FUNCTION "FRK_Release_DeclarationUnit" : Void
{ S7_Optimized_Access := 'TRUE' }
VERSION : 0.1
VAR_IN_OUT
    Unit : "FRK_Unit";
    Hal : "ST_DeclarationUnitHal";
END_VAR
BEGIN
    "FRK_UnitSetPermit"(Unit := #Unit, Ok := #Hal.Cell.Clamp.Permit, Diag := #Hal.Cell.Clamp.Diag);
END_FUNCTION
// Generated frame v0.24; change the declaration, then regenerate.
FUNCTION_BLOCK "FB_DeclarationUnit"
{ S7_Optimized_Access := 'TRUE' }
VERSION : 0.1
VAR_INPUT
    Execute {ExternalWritable := 'False'} : Bool;
    Abort {ExternalWritable := 'False'} : Bool;
    Command {ExternalWritable := 'False'} : DInt;
    ParCmd {ExternalWritable := 'False'} : "ST_DeclarationParCmd";
    ParentIndex {ExternalAccessible := 'False'; ExternalVisible := 'False'; ExternalWritable := 'False'} : DInt;
    Startup {ExternalAccessible := 'False'; ExternalVisible := 'False'; ExternalWritable := 'False'} : Bool;
END_VAR
VAR_OUTPUT
    Busy {ExternalWritable := 'False'} : Bool;
    Done {ExternalWritable := 'False'} : Bool;
    Error {ExternalWritable := 'False'} : Bool;
    Aborted {ExternalWritable := 'False'} : Bool;
    Held {ExternalWritable := 'False'} : Bool;
    ErrorID {ExternalWritable := 'False'} : DWord;
    Timing {ExternalWritable := 'False'} : "ST_ModuleTiming";
    OutCmd {ExternalWritable := 'False'} : "ST_DeclarationOutCmd";
END_VAR
VAR_IN_OUT
    Hal : "ST_DeclarationUnitHal";
END_VAR
VAR
    OutImm {ExternalWritable := 'False'} : "ST_UnitProbeImm";
    Status {ExternalWritable := 'False'} : "ST_ModuleStatus";
    Core {ExternalAccessible := 'False'; ExternalVisible := 'False'; ExternalWritable := 'False'} : "FRK_Core";
    Nameplate {ExternalWritable := 'False'} : "ST_Nameplate";
    EngineeringSlots {ExternalAccessible := 'False'; ExternalVisible := 'False'; ExternalWritable := 'False'} : Array[1..1] of Int;
    RunStyle {ExternalWritable := 'False'} : DInt;
    SupportedRunStylesPublished {ExternalWritable := 'False'} : Array[0..2] of Bool;
    HostEvents {ExternalWritable := 'False'} : "FRK_HostEvents";
    HostSeenSequence {ExternalAccessible := 'False'; ExternalVisible := 'False'; ExternalWritable := 'False'} : UDInt;
    HostDoneSeen {ExternalAccessible := 'False'; ExternalVisible := 'False'; ExternalWritable := 'False'} : Bool;
    SystemHealth {ExternalWritable := 'False'} : "ST_SystemHealthStatus";
    HealthBook {ExternalAccessible := 'False'; ExternalVisible := 'False'; ExternalWritable := 'False'} : "FRK_HealthBook";
    HealthConfig {ExternalAccessible := 'False'; ExternalVisible := 'False'; ExternalWritable := 'False'} : "ST_SystemHealthParCfg";
    SignalTower {ExternalWritable := 'False'} : "ST_SignalTowerOut";
    TowerBook {ExternalAccessible := 'False'; ExternalVisible := 'False'; ExternalWritable := 'False'} : "FRK_TowerBook";
    TowerConfig {ExternalAccessible := 'False'; ExternalVisible := 'False'; ExternalWritable := 'False'} : "ST_SignalTowerParCfg";
    ParCfg {ExternalWritable := 'False'} : "ST_ProductionUnitParCfg";
    LatchedParCmd {ExternalAccessible := 'False'; ExternalVisible := 'False'; ExternalWritable := 'False'} : "ST_DeclarationParCmd";
    StateFlags {ExternalWritable := 'False'} : Array[1..12] of "ST_StateFlag";
    StateFlagCount {ExternalWritable := 'False'} : Int;
    StateTouched {ExternalAccessible := 'False'; ExternalVisible := 'False'; ExternalWritable := 'False'} : Array[1..12] of Bool;
    Device {ExternalAccessible := 'False'; ExternalVisible := 'False'; ExternalWritable := 'False'} : "ST_UnitProbeDevice";
    StationCfg {ExternalWritable := 'False'} : "ST_UnitProbeStationCfg";
    ConfigStageParCfg {ExternalAccessible := 'False'; ExternalVisible := 'False'; ExternalWritable := 'False'} : "ST_ProductionUnitParCfg";
    ConfigDefaultParCfg {ExternalAccessible := 'False'; ExternalVisible := 'False'; ExternalWritable := 'False'} : "ST_ProductionUnitParCfg";
    ConfigStageStationCfg {ExternalAccessible := 'False'; ExternalVisible := 'False'; ExternalWritable := 'False'} : "ST_UnitProbeStationCfg";
    ConfigDefaultStationCfg {ExternalAccessible := 'False'; ExternalVisible := 'False'; ExternalWritable := 'False'} : "ST_UnitProbeStationCfg";
    ConfigStaged {ExternalAccessible := 'False'; ExternalVisible := 'False'; ExternalWritable := 'False'} : Bool;
    ConfigPersist {ExternalWritable := 'False'} : "ST_ConfigPersistStatus";
    Model {ExternalWritable := 'False'} : "ST_ModelId";
    AvailableModelCount {ExternalWritable := 'False'} : Int;
    AvailableModels {ExternalWritable := 'False'} : Array[1..3] of "ST_ModelId";
    ModelCapacity {ExternalWritable := 'False'} : Int;
    ModelGenerationSeen {ExternalAccessible := 'False'; ExternalVisible := 'False'; ExternalWritable := 'False'} : UDInt;
    ConfigSets {ExternalWritable := 'False'} : Array[1..4] of "ST_ConfigSetInfo";
    ConfigSetCount {ExternalWritable := 'False'} : Int;
    ConfigSetDocument {ExternalWritable := 'False'} : WString[480];
    ConfigSetDocumentLine {ExternalWritable := 'False'} : Int;
    ConfigSetDocumentLines {ExternalWritable := 'False'} : Int;
    SequenceViewEnabled {ExternalWritable := 'False'} : Bool;
    SequenceStepCount {ExternalWritable := 'False'} : Int;
    SequenceAnnotationCount {ExternalWritable := 'False'} : Int;
    Pending {ExternalWritable := 'False'} : "ST_Diagnostic";
    CurrentStep {ExternalWritable := 'False'} : "ST_StepRecord";
    CurrentStepElapsed {ExternalWritable := 'False'} : Time;
    CurrentStepTimedOut {ExternalWritable := 'False'} : Bool;
    SequenceSteps {ExternalWritable := 'False'} : Array[1..8] of "ST_SequenceStep";
    ActiveSteps {ExternalWritable := 'False'} : Array[0..0] of "ST_SequenceCursor";
    SequenceAnnotations {ExternalWritable := 'False'} : Array[1..4] of "ST_SequenceAnnotation";
    SequenceStepDef {ExternalAccessible := 'False'; ExternalVisible := 'False'; ExternalWritable := 'False'} : Array[1..8] of "ST_SequenceStepDef";
    Profiler {ExternalWritable := 'False'} : "FRK_Profiler_DeclarationUnit";
    Starved {ExternalWritable := 'False'} : Bool;
    Blocked {ExternalWritable := 'False'} : Bool;
    ProductionBook {ExternalAccessible := 'False'; ExternalVisible := 'False'; ExternalWritable := 'False'} : "FRK_Production";
    MachineState {ExternalWritable := 'False'} : DInt;
    Oee {ExternalWritable := 'False'} : "ST_Oee";
    OeeTrend {ExternalWritable := 'False'} : Array[1..60] of "ST_OeeSample";
    OeeTrendHead {ExternalWritable := 'False'} : Int;
    Unit {ExternalAccessible := 'False'; ExternalVisible := 'False'; ExternalWritable := 'False'} : "FRK_Unit";
    HmiRequest : "ST_HmiRequest";
    ModePolicy {ExternalAccessible := 'False'; ExternalVisible := 'False'; ExternalWritable := 'False'} : Array[0..6] of "ST_ModePolicy";
    Access {ExternalWritable := 'False'} : "FRK_Access";
    HmiResponse {ExternalWritable := 'False'} : "ST_HmiResponse";
    ConfigRev {ExternalWritable := 'False'} : UDInt;
    ConfigCursor {ExternalAccessible := 'False'; ExternalVisible := 'False'; ExternalWritable := 'False'} : "FRK_ConfigCursor";
    Part {ExternalWritable := 'False'} : "ST_PartContext";
    Decision {ExternalWritable := 'False'} : "ST_DecisionRequest";
    DecisionAnswer {ExternalWritable := 'False'} : Int;
    History {ExternalWritable := 'False'} : Array[1..16] of "ST_Diagnostic";
    HistoryHead {ExternalWritable := 'False'} : Int;
    AlarmLog {ExternalWritable := 'False'} : "FRK_AlarmLog";
    ModeActivePublished {ExternalWritable := 'False'} : DInt;
    RunningPublished {ExternalWritable := 'False'} : Bool;
    StopPendingPublished {ExternalWritable := 'False'} : Bool;
    SupportedModesPublished {ExternalWritable := 'False'} : Array[0..6] of Bool;
    GoodCount {ExternalWritable := 'False'} : UDInt;
    NokCount {ExternalWritable := 'False'} : UDInt;
    ReworkCount {ExternalWritable := 'False'} : UDInt;
    NokReason {ExternalWritable := 'False'} : DInt;
    Cell {ExternalWritable := 'False'} : "FB_DeclarationCell";
    Satellite {ExternalWritable := 'False'} : "FB_SatelliteUnit";
END_VAR
VAR_TEMP
    InstancePath : WString[254];
    RouteMatched : Bool;
    ManualMatched : Bool;
    ConfigRootIndex : Int;
    HealthResult : Bool;
END_VAR
VAR CONSTANT
    EXEC_READY : DInt := 0;
    MODULE_TIER : DInt := 1;
END_VAR
BEGIN
    // ---- GENERATED: setup
    IF #Startup OR NOT #Core.Named THEN
        #InstancePath := GetInstancePath(SIZE := 0);
        "FRK_SetIdentity"(Core := #Core, Status := #Status, InstancePath := #InstancePath,
            ModuleType := 1, TypeId := 1, Capabilities := DWORD#16#00000000, ParentIndex := #ParentIndex, TypeKey := 'Fraktal.Declaration.Unit');
        IF #Core.RegIndex = 1 THEN
            #Nameplate.ProductUri := WSTRING#'urn:fraktal:tia:operations:station-a';
            #Nameplate.ManufacturerName := 'Fraktal';
            #Nameplate.ProductDesignation := 'Isolated operations fixture';
        END_IF;
    END_IF;
    IF #Startup THEN "FRK_CfgRestore_DeclarationUnit"(Core := #Core, Status := #Status, ParCfg := #ParCfg, StationCfg := #StationCfg, ConfigStageParCfg := #ConfigStageParCfg, ConfigDefaultParCfg := #ConfigDefaultParCfg, ConfigStageStationCfg := #ConfigStageStationCfg, ConfigDefaultStationCfg := #ConfigDefaultStationCfg); END_IF;
    #ConfigRootIndex := "FRK_ConfigRoot"(RegIndex := #Core.RegIndex);
    "FRK_StateSweep"(Flags := #StateFlags, Count := #StateFlagCount, Touched := #StateTouched, Startup := #Startup);
    IF #Startup OR #ConfigRev = 0 THEN #ConfigRev := "FRK_ConfigRevision"(Previous := #ConfigRev); END_IF;
    #SupportedModesPublished[0] := TRUE;
    #SupportedModesPublished[1] := TRUE;
    #SupportedModesPublished[2] := TRUE;
    #SupportedModesPublished[3] := TRUE;
    #SupportedModesPublished[4] := FALSE;
    #SupportedModesPublished[5] := FALSE;
    #SupportedModesPublished[6] := FALSE;
    "FRK_UnitPrepare"(Core := #Core, Unit := #Unit, Policy := #ModePolicy, Request := #HmiRequest, Response := #HmiResponse, Startup := #Startup, InitialMode := 1);
    "FRK_AlarmBegin"(AlarmLog := #AlarmLog, Startup := #Startup);
    "FRK_AlarmHistoryBoot"(AlarmLog := #AlarmLog, Startup := #Startup, Scope := #Status.Name);
    "FRK_AlarmRecoveryBoot"(AlarmLog := #AlarmLog, Startup := #Startup, Scope := #Status.Name);
    "FRK_AlarmRecoveryTick"(AlarmLog := #AlarmLog);
    "FRK_AccessPolicyBoot"(Access := #Access, Startup := #Startup, Root := #Core.ParentIndex = 0, Scope := #Status.Name);
    "FRK_ClassBoot"(Access := #Access, Startup := #Startup, Root := #Core.ParentIndex = 0, Scope := #Status.Name);
    "FRK_AccessCyclic"(Access := #Access, Startup := #Startup, SourcePath := STRING_TO_WSTRING(#Status.Name), AlarmLog := #AlarmLog, Revision := #ConfigRev);
    "FRK_UnitMailbox"(Core := #Core, Unit := #Unit, Status := #Status, Policy := #ModePolicy, Access := #Access, Request := #HmiRequest, Response := #HmiResponse, Supported := #SupportedModesPublished);
    "FRK_ConfigStatus"(RootIndex := #ConfigRootIndex, Scope := #Status.Name, PolicyLost := (#Access.PolicyLost OR #Access.ClassesLost), UsersLost := "FRK_AccessStorage".UsersLost, Persist := #ConfigPersist, AlarmLog := #AlarmLog);
    #Unit.ConfigEnabled := #Core.ParentIndex = 0;
    #Unit.ConfigSetsEnabled := TRUE AND #Core.ParentIndex = 0;
    #Unit.ModelEnabled := #AvailableModelCount > 0;
    #Unit.ConfigBlocked := #ConfigPersist.RestoreLost AND NOT #ConfigPersist.RestoreAcknowledged AND #ConfigPersist.RestorePolicy = 1;
    #Unit.ConfigBlocked := #Unit.ConfigBlocked OR (#Access.PolicyLost OR #Access.ClassesLost);
    // ---- GENERATED: begin
    "FRK_Begin"(Core := #Core, Status := #Status, Execute := #Unit.RunReq, Abort := (#Abort OR #Unit.AbortReq), Command := 1);
    IF #Core.EvCommandStart THEN
        #LatchedParCmd := #ParCmd;
        CASE #Core.Command OF
            1: "FRK_UnitRunStart"(Core := #Core, Status := #Status, Timeout := #ParCfg.Timeout, Label := 'Run');
            ELSE "FRK_Start"(Core := #Core, Status := #Status, Supported := FALSE, Timeout := T#0ms, Label := '');
        END_CASE;
    END_IF;
    IF #Core.EvCommandStart THEN
    // ---- AUTHORED: CommandStart
    #Device.Received := "FRK_PartReceived"(Core := #Core, Unit := #Unit, Status := #Status, Part := #Part, AlarmLog := #AlarmLog);
    IF #Device.Received THEN
        "FRK_PartStarted"(Unit := #Unit, Status := #Status, Part := #Part, AlarmLog := #AlarmLog);
    END_IF;
    // ---- GENERATED: reaction end
    END_IF;
    IF #Core.EvCommandStart AND #Unit.Mode = 3 THEN
        "FRK_HostEmit"(Kind := 5, Scope := #Status.Name, PartUid := '', Subject := 'Model', Value := #Model.ModelCode, Verdict := 0, Reason := 0);
    END_IF;
    // ---- AUTHORED: cyclic management
    IF #Hal.Cell.Clamp.BackgroundFault THEN
        "FRK_Fault"(Core := #Core, Status := #Status, ReasonCode := 2901, Description := WSTRING#'test.unit.condition');
    END_IF;
    // ---- GENERATED: end management
    "FRK_Release_DeclarationUnit"(Unit := #Unit, Hal := #Hal);
    IF #Core.RegIndex > 0 THEN "FRK_Registry".Rows[#Core.RegIndex].AlarmBlocking := #AlarmLog.Blocking; END_IF;
    #Unit.AlarmBlocking := "FRK_AlarmTreeBlocking"(Owner := #Core.RegIndex) OR "FRK_AlarmRecoveryTreeBlocking"(Scope := #Status.Name);
    "FRK_UnitConsume"(Core := #Core, Unit := #Unit, Status := #Status, Policy := #ModePolicy, Access := #Access, Response := #HmiResponse, Supported := #SupportedModesPublished);
    "FRK_UnitMode"(Core := #Core, Unit := #Unit);
    #SupportedRunStylesPublished[0] := TRUE;
    #SupportedRunStylesPublished[1] := FALSE;
    #SupportedRunStylesPublished[2] := FALSE;
    "FRK_RunStylePrepare"(Owner := #Core.RegIndex, Startup := #Startup OR #Core.EvModeChanged OR #Unit.EvReset, Exec := #Core.Exec, Access := #Access, Supported := #SupportedRunStylesPublished);
    "FRK_RunStyleRequest"(Owner := #Core.RegIndex, Scope := #Status.Name, Exec := #Core.Exec, Supported := #SupportedRunStylesPublished, Unit := #Unit, Access := #Access, Response := #HmiResponse);
    "FRK_AlarmShelfRequest"(Scope := #Status.Name, Unit := #Unit, Access := #Access, Response := #HmiResponse, AlarmLog := #AlarmLog);
    #TowerConfig := "FRK_TowerDefaults".Config;
    "FRK_TowerRequest"(Scope := #Status.Name, Core := #Core, Unit := #Unit, Access := #Access, Response := #HmiResponse, Book := #TowerBook, ParCfg := #TowerConfig);
    "FRK_ProductionRequest"(Unit := #Unit, Access := #Access, Response := #HmiResponse, Book := #ProductionBook, Oee := #Oee, Trend := #OeeTrend, AlarmLog := #AlarmLog, Scope := #Status.Name);
    IF #Core.EvModeExit THEN
    // ---- AUTHORED: ModeExit
    #Device.ExitCalls := #Device.ExitCalls + 1;
    IF #Hal.Cell.Clamp.ExitHold THEN #Core.HookResult := 1; ELSE #Core.HookResult := 0; END_IF;
    // ---- GENERATED: reaction end
    END_IF;
    "FRK_UnitModeResolve"(Core := #Core, Unit := #Unit, Status := #Status, Policy := #ModePolicy, Timeout := #ParCfg.Timeout);
    IF #Core.EvModeChanged THEN
    // ---- AUTHORED: ModeChanged
    #Device.Changes := #Device.Changes + 1;
    // ---- GENERATED: reaction end
    END_IF;
    IF #Core.EvModeChanged THEN
        "FRK_HostEmit"(Kind := 9, Scope := #Status.Name, PartUid := '', Subject := 'Mode', Value := DINT_TO_STRING(#Unit.Mode), Verdict := 0, Reason := 0);
    END_IF;
    "FRK_SeqViewBegin"(Owner := #Core.RegIndex, Clear := #Startup OR #Core.EvModeChanged, ResetErrors := #Unit.EvReset, Enabled := #SequenceViewEnabled);
    "FRK_SeqProfilePrepare"(Owner := #Core.RegIndex, Run := #Core.Exec = 1 AND #Unit.Mode = 0, Withdraw := #Startup OR #Core.EvModeChanged);
    "FRK_DecisionCyclic"(Owner := #Core.RegIndex, Busy := #Core.Exec = 1, Reset := #Startup OR #Unit.EvReset OR #Core.EvModeChanged, AlarmLog := #AlarmLog);
    "FRK_UnitFollow"(Core := #Core, Unit := #Unit, Status := #Status, Policy := #ModePolicy, Access := #Access, Supported := #SupportedModesPublished);
    IF #Unit.RequestPending AND (#Unit.Request.Kind = 11 OR #Unit.Request.Kind = 16) THEN
        #ManualMatched := FALSE;
        #RouteMatched := "FRK_Route_DeclarationCell"(Module := #Cell, Hal := #Hal.Cell, Request := #Unit.Request, Report := #HmiResponse.Report);
        #ManualMatched := #ManualMatched OR #RouteMatched;
        #RouteMatched := "FRK_Route_SatelliteUnit"(Module := #Satellite, Hal := #Hal.Satellite, Request := #Unit.Request, Report := #HmiResponse.Report);
        #ManualMatched := #ManualMatched OR #RouteMatched;
        IF NOT #ManualMatched THEN
            "FRK_ReleaseReason"(Report := #HmiResponse.Report, Description := WSTRING#'std.error.unsupportedHmiRequest', Reason := 2008, Path := #Unit.Request.TargetPath, Kind := 4);
        END_IF;
        #HmiResponse.Accepted := #Unit.Request.Kind = 16 OR #HmiResponse.Report.Released;
        IF #Unit.Request.Kind = 11 THEN
            IF #HmiResponse.Accepted THEN #HmiResponse.Diagnostic := WSTRING#'std.audit.manualCommandAccepted'; ELSE #HmiResponse.Diagnostic := WSTRING#'std.audit.manualCommandRejected'; END_IF;
        END_IF;
    END_IF;
    IF #Unit.EvReset THEN "FRK_AlarmOperatorReset"(AlarmLog := #AlarmLog); END_IF;
    IF #Unit.EvReset THEN
    // ---- AUTHORED: OperatorReset
    #Device.Resets := #Device.Resets + 1;
    // ---- GENERATED: reset reaction end
    END_IF;
    IF #Core.ReleasePending OR #Unit.ReleaseChildren THEN
        "FRK_ReleaseCommand"(Core := #Cell.Core, Execute := #Cell.Execute);
        "FRK_ReleaseCommand"(Core := #Satellite.Core, Execute := #Satellite.Execute);
    END_IF;
    // ---- GENERATED: child call
    #Cell(ParentIndex := #Core.RegIndex, Startup := #Startup, Hal := #Hal.Cell);
    "FRK_ManualFinish"(Core := #Cell.Core, Execute := #Cell.Execute, ManualOwned := #Cell.ManualOwned);
    "FRK_UnitCascade"(ParentUnit := #Unit, Core := #Satellite.Core, Unit := #Satellite.Unit, Status := #Satellite.Status, Policy := #Satellite.ModePolicy, Access := #Satellite.Access, Supported := #Satellite.SupportedModesPublished, AlarmLog := #AlarmLog);
    // ---- GENERATED: child call
    #Satellite(ParentIndex := #Core.RegIndex, Startup := #Startup, Hal := #Hal.Satellite);
    #Unit.CascadePending := FALSE;
    "FRK_ConfigScratch".AccessRejected := FALSE;
    "FRK_CfgModelOperation_DeclarationUnit"(Core := #Core, Status := #Status, ParCfg := #ParCfg, Access := #Access, Unit := #Unit, HmiResponse := #HmiResponse, AlarmLog := #AlarmLog, ConfigPersist := #ConfigPersist, ConfigRev := #ConfigRev, AvailableModelCount := #AvailableModelCount, ModelCapacity := #ModelCapacity, ModelGenerationSeen := #ModelGenerationSeen, AvailableModels := #AvailableModels, StationCfg := #StationCfg, ConfigStageParCfg := #ConfigStageParCfg, ConfigStageStationCfg := #ConfigStageStationCfg, Cell := #Cell, Satellite := #Satellite);
    "FRK_CfgOperation_DeclarationUnit"(Core := #Core, Status := #Status, OutImm := #OutImm, ParCfg := #ParCfg, ModePolicy := #ModePolicy, Access := #Access, Unit := #Unit, HmiResponse := #HmiResponse, AlarmLog := #AlarmLog, ConfigPersist := #ConfigPersist, ConfigCursor := #ConfigCursor, ConfigRev := #ConfigRev, Model := #Model, AvailableModelCount := #AvailableModelCount, ConfigStaged := #ConfigStaged, ModelCapacity := #ModelCapacity, SequenceStepDef := #SequenceStepDef, SequenceStepCount := #SequenceStepCount, SupportedModesPublished := #SupportedModesPublished, StationCfg := #StationCfg, ConfigStageParCfg := #ConfigStageParCfg, ConfigDefaultParCfg := #ConfigDefaultParCfg, Cell := #Cell, Satellite := #Satellite);
    "FRK_CfgSetOperation_DeclarationUnit"(Core := #Core, Status := #Status, ParCfg := #ParCfg, ModePolicy := #ModePolicy, Access := #Access, Unit := #Unit, HmiResponse := #HmiResponse, ConfigPersist := #ConfigPersist, ConfigRev := #ConfigRev, Model := #Model, AvailableModelCount := #AvailableModelCount, ConfigSets := #ConfigSets, ConfigSetCount := #ConfigSetCount, ConfigSetDocument := #ConfigSetDocument, ConfigSetDocumentLine := #ConfigSetDocumentLine, ConfigSetDocumentLines := #ConfigSetDocumentLines, SupportedModesPublished := #SupportedModesPublished, StationCfg := #StationCfg, ConfigStageParCfg := #ConfigStageParCfg, ConfigStageStationCfg := #ConfigStageStationCfg, Cell := #Cell, Satellite := #Satellite, Startup := #Startup);
    IF #Unit.RequestPending AND #Core.ParentIndex = 0 THEN "FRK_SetResult"(Request := #Unit.Request, Response := #HmiResponse, Persist := #ConfigPersist, AlarmLog := #AlarmLog, Scope := #Status.Name, RootIndex := #ConfigRootIndex); END_IF;
    "FRK_ConfigAccessRefusal"(Unit := #Unit, Access := #Access, Response := #HmiResponse, Persist := #ConfigPersist, AlarmLog := #AlarmLog);
    "FRK_ConfigStatus"(RootIndex := #ConfigRootIndex, Scope := #Status.Name, PolicyLost := (#Access.PolicyLost OR #Access.ClassesLost), UsersLost := "FRK_AccessStorage".UsersLost, Persist := #ConfigPersist, AlarmLog := #AlarmLog);
    "FRK_RouteAbort"(Core := #Core, Abort := (#Abort OR #Unit.AbortReq));
    IF #Core.EvAbort THEN
        "FRK_PartAborted"(Core := #Core, Unit := #Unit, Status := #Status, Part := #Part, AlarmLog := #AlarmLog);
    END_IF;
    "FRK_SeqLifecycleUpdate"(Owner := #Core.RegIndex, Exec := #Core.Exec, Restart := #Startup OR #Core.EvModeChanged OR #Core.EvAbortInError);
    "FRK_DiagComposite"(Core := #Core, Status := #Status, AdoptErrors := FALSE);
    IF #Core.Dispatch AND #Core.RegIndex > 0 AND NOT "FRK_Registry".Fault THEN
    // ---- AUTHORED: dispatch
    IF #Hal.Cell.Clamp.Finish THEN
        #Device.Processed := FALSE;
        IF #Unit.CarrierIndex = 0 THEN
            #Device.Processed := TRUE;
        ELSE
            #Device.Processed := "FRK_PartProcessed"(Core := #Core, Unit := #Unit, Status := #Status, Part := #Part, AlarmLog := #AlarmLog, Verdict := #Hal.Cell.Clamp.Verdict, Reason := #Hal.Cell.Clamp.Diag.ReasonCode);
        END_IF;
        IF #Device.Processed THEN
            #Device.Cycles := #Device.Cycles + 1;
            IF #Unit.StopReq THEN
                "FRK_Complete"(Core := #Core, Status := #Status);
            ELSE
                #Device.Received := "FRK_PartReceived"(Core := #Core, Unit := #Unit, Status := #Status, Part := #Part, AlarmLog := #AlarmLog);
                IF #Device.Received THEN
                    "FRK_PartStarted"(Unit := #Unit, Status := #Status, Part := #Part, AlarmLog := #AlarmLog);
                END_IF;
            END_IF;
        END_IF;
    END_IF;
    // ---- GENERATED: end dispatch
    END_IF;
    "FRK_SeqViewEnd"(Owner := #Core.RegIndex, Revision := #ConfigRev, Fallback := #ParCfg.Timeout);
    "FRK_SeqViewDiagnostic"(Owner := #Core.RegIndex, Core := #Core, Status := #Status, Pending := #Pending);
    CASE #Core.RegIndex OF
        1:
            #SequenceStepDef := "FRK_Views".V001.Defs;
            #SequenceSteps := "FRK_Views".V001.Rows;
            #ActiveSteps := "FRK_Views".V001.Cursors;
            #SequenceAnnotations := "FRK_Views".V001.Notes;
            #SequenceStepCount := "FRK_Views".V001.Count;
            #SequenceAnnotationCount := "FRK_Views".V001.NoteCount;
            #CurrentStep := "FRK_Views".V001.Current;
            #CurrentStepElapsed := "FRK_Views".V001.Cursors[0].Elapsed;
            #CurrentStepTimedOut := "FRK_Views".V001.Cursors[0].TimedOut;
        13:
            #SequenceStepDef := "FRK_Views".V013.Defs;
            #SequenceSteps := "FRK_Views".V013.Rows;
            #ActiveSteps := "FRK_Views".V013.Cursors;
            #SequenceAnnotations := "FRK_Views".V013.Notes;
            #SequenceStepCount := "FRK_Views".V013.Count;
            #SequenceAnnotationCount := "FRK_Views".V013.NoteCount;
            #CurrentStep := "FRK_Views".V013.Current;
            #CurrentStepElapsed := "FRK_Views".V013.Cursors[0].Elapsed;
            #CurrentStepTimedOut := "FRK_Views".V013.Cursors[0].TimedOut;
        ELSE #SequenceViewEnabled := FALSE;
    END_CASE;
    "FRK_End"(Core := #Core, Status := #Status,
        Busy => #Busy, Done => #Done, Error => #Error, Aborted => #Aborted, Held => #Held, ErrorID => #ErrorID, Timing => #Timing);
    "FRK_SeqLifecycleUpdate"(Owner := #Core.RegIndex, Exec := #Core.Exec, Restart := FALSE);
    IF #Core.Exec = 3 OR #Core.Exec = 4 THEN
        "FRK_SeqProfilePrepare"(Owner := #Core.RegIndex, Run := FALSE, Withdraw := TRUE);
    END_IF;
    "FRK_SeqProfileEnd"(Owner := #Core.RegIndex, StepNo := #CurrentStep.StepNo, Expected := #CurrentStep.ExpectedTime, NowMs := "FRK_Clock".NowMs);
    CASE #Core.RegIndex OF
        1:
            #Profiler.LastCycle.CycleNo := "FRK_Profiles".P001.Book.Last.CycleNo;
            #Profiler.LastCycle.Started := "FRK_Profiles".P001.Book.Last.Started;
            #Profiler.LastCycle.StartedTimeSynchronized := "FRK_Profiles".P001.Book.Last.StartedTimeSynchronized;
            #Profiler.LastCycle.Total := "FRK_Profiles".P001.Book.Last.Total;
            #Profiler.LastCycle.WorkTime := "FRK_Profiles".P001.Book.Last.WorkTime;
            #Profiler.LastCycle.WaitTime := "FRK_Profiles".P001.Book.Last.WaitTime;
            #Profiler.LastCycle.ByClass := "FRK_Profiles".P001.Book.Last.ByClass;
            #Profiler.LastCycle.NSteps := "FRK_Profiles".P001.Book.LastNSteps;
            #Profiler.LastCycle.Truncated := "FRK_Profiles".P001.Book.LastTruncated;
            #Profiler.LastCycle.Steps := "FRK_Profiles".P001.LastSteps;
            #Profiler.StepStats := "FRK_Profiles".P001.Stats;
            #Profiler.StatsTruncated := "FRK_Profiles".P001.Book.StatsTruncated;
            #Profiler.LastCycleTime := "FRK_Profiles".P001.Book.LastCycleTime;
            #Profiler.MinCycleTime := "FRK_Profiles".P001.Book.MinCycleTime;
            #Profiler.History := "FRK_Profiles".P001.History;
            #Profiler.HistoryHead := "FRK_Profiles".P001.Book.Head;
        13:
            #Profiler.LastCycle.CycleNo := "FRK_Profiles".P013.Book.Last.CycleNo;
            #Profiler.LastCycle.Started := "FRK_Profiles".P013.Book.Last.Started;
            #Profiler.LastCycle.StartedTimeSynchronized := "FRK_Profiles".P013.Book.Last.StartedTimeSynchronized;
            #Profiler.LastCycle.Total := "FRK_Profiles".P013.Book.Last.Total;
            #Profiler.LastCycle.WorkTime := "FRK_Profiles".P013.Book.Last.WorkTime;
            #Profiler.LastCycle.WaitTime := "FRK_Profiles".P013.Book.Last.WaitTime;
            #Profiler.LastCycle.ByClass := "FRK_Profiles".P013.Book.Last.ByClass;
            #Profiler.LastCycle.NSteps := "FRK_Profiles".P013.Book.LastNSteps;
            #Profiler.LastCycle.Truncated := "FRK_Profiles".P013.Book.LastTruncated;
            #Profiler.LastCycle.Steps := "FRK_Profiles".P013.LastSteps;
            #Profiler.StepStats := "FRK_Profiles".P013.Stats;
            #Profiler.StatsTruncated := "FRK_Profiles".P013.Book.StatsTruncated;
            #Profiler.LastCycleTime := "FRK_Profiles".P013.Book.LastCycleTime;
            #Profiler.MinCycleTime := "FRK_Profiles".P013.Book.MinCycleTime;
            #Profiler.History := "FRK_Profiles".P013.History;
            #Profiler.HistoryHead := "FRK_Profiles".P013.Book.Head;
        ELSE RETURN;
    END_CASE;
    #Starved := #Core.Exec = 1 AND #Unit.Mode = 0 AND #CurrentStep.TimeClass = 1;
    #Blocked := #Core.Exec = 1 AND #Unit.Mode = 0 AND #CurrentStep.TimeClass = 2;
    "FRK_DecisionCyclic"(Owner := #Core.RegIndex, Busy := #Core.Exec = 1, Reset := #Startup OR #Unit.EvReset OR #Core.EvModeChanged, AlarmLog := #AlarmLog);
    "FRK_DecisionPublish"(Owner := #Core.RegIndex, Decision := #Decision, DecisionAnswer := #DecisionAnswer);
    IF NOT #Unit.EvReset THEN
        "FRK_AlarmCapture"(AlarmLog := #AlarmLog, Core := #Core, Status := #Status);
        "FRK_Capture_DeclarationCell"(Module := #Cell, AlarmLog := #AlarmLog);
        "FRK_AlarmEnd"(AlarmLog := #AlarmLog);
    END_IF;
    IF #Core.RegIndex > 0 THEN "FRK_Registry".Rows[#Core.RegIndex].AlarmBlocking := #AlarmLog.Blocking; END_IF;
    #Unit.AlarmBlocking := "FRK_AlarmTreeBlocking"(Owner := #Core.RegIndex) OR "FRK_AlarmRecoveryTreeBlocking"(Scope := #Status.Name);
    "FRK_ClassOperation"(Access := #Access, Unit := #Unit, Response := #HmiResponse, Scope := #Status.Name);
    "FRK_AccessPersist"(Access := #Access, Unit := #Unit, Response := #HmiResponse, SourcePath := STRING_TO_WSTRING(#Status.Name), AlarmLog := #AlarmLog);
    IF #Core.ParentIndex = 0 THEN "FRK_EngineeringTick"(Scope := #Status.Name, Slots := #EngineeringSlots, AlarmLog := #AlarmLog); END_IF;
    #HealthConfig := "FRK_HealthDefaults".Config;
    #HealthResult := "FRK_HealthCyclic"(Configured := TRUE, Scope := #Status.Name, Input := "FRK_HealthProbe".Input, ParCfg := #HealthConfig, Status := #SystemHealth, Book := #HealthBook, AlarmLog := #AlarmLog);
    IF #Startup THEN #ProductionBook := "FRK_ProductionDefaults".Book; #Oee := "FRK_ProductionDefaults".Oee; END_IF;
    #MachineState := "FRK_MachineState"(Exec := #Core.Exec, Mode := #Unit.Mode, Blocking := #Unit.AlarmBlocking, Starved := #Starved, Blocked := #Blocked, StopRequested := #Unit.StopReq);
    "FRK_OeeTick"(NowMs := "FRK_Clock".NowMs, Exec := #Core.Exec, Blocking := #Unit.AlarmBlocking, Good := #Unit.Good, Nok := #Unit.Nok, IdealCycleMs := #ParCfg.IdealCycleMs, Book := #ProductionBook, Oee := #Oee, Trend := #OeeTrend);
    #OeeTrendHead := #ProductionBook.TrendHead;
    IF "FRK_WorkDegradation"(CycleNo := #Profiler.LastCycle.CycleNo, WorkMs := TIME_TO_UDINT(#Profiler.LastCycle.WorkTime), BaselineMs := #ParCfg.BaselineMs, BandPercent := #StationCfg.DegradationPercent, Book := #ProductionBook) THEN
        "FRK_AlarmMessage"(AlarmLog := #AlarmLog, Reason := 2007, Description := WSTRING#'std.maintenance.cycleTimeDegraded', SourcePath := STRING_TO_WSTRING(#Status.Name));
    END_IF;
    IF #Startup THEN #TowerBook.TestActive := FALSE; END_IF;
    "FRK_TowerFrame"(MachineState := #MachineState, OperatorActionRequired := #Decision.Prompt <> WSTRING#'' OR "FRK_Registry".Rows[#Core.RegIndex].StepWait, ParCfg := #TowerConfig, Book := #TowerBook, AlarmLog := #AlarmLog, Status := #SignalTower);
    IF #Core.Exec = 2 AND NOT #HostDoneSeen AND #Unit.Mode = 3 THEN
        "FRK_HostEmit"(Kind := 6, Scope := #Status.Name, PartUid := '', Subject := 'Model', Value := #Model.ModelCode, Verdict := 0, Reason := 0);
    END_IF;
    #HostDoneSeen := #Core.Exec = 2;
    "FRK_HostMirror"(Scope := #Status.Name, Startup := #Startup, Seen := #HostSeenSequence, View := #HostEvents);
    "FRK_AccessFinish"(Access := #Access, Unit := #Unit, Response := #HmiResponse, SourcePath := STRING_TO_WSTRING(#Status.Name), AlarmLog := #AlarmLog, Revision := #ConfigRev);
    "FRK_UnitFinish"(Core := #Core, Unit := #Unit, Response := #HmiResponse, Status := #Status, Part := #Part, AlarmLog := #AlarmLog, History := #History, Head := #HistoryHead);
    #ModeActivePublished := #Unit.Mode;
    #RunningPublished := #Core.Exec = 1;
    #StopPendingPublished := #Unit.StopReq AND #Core.Exec = 1;
    #GoodCount := #Unit.Good;
    #NokCount := #Unit.Nok;
    #ReworkCount := #Unit.Rework;
    #NokReason := #Unit.NokReason;
    IF #Core.RegIndex > 0 THEN #RunStyle := "FRK_Registry".Rows[#Core.RegIndex].RunStyle; END_IF;
    // ---- AUTHORED: unconditional cyclic/derived data
    #OutImm.Cycles := #Device.Cycles;
    #OutImm.ExitCalls := #Device.ExitCalls;
    #OutImm.Changes := #Device.Changes;
    #OutImm.Resets := #Device.Resets;
    #OutImm.AtHome := "FRK_State"(Idx := 1, Key := 'project.state.atHome', Ok := #Hal.Cell.Clamp.Sample = 0, Flags := #StateFlags, Count := #StateFlagCount, Touched := #StateTouched);
    // ---- GENERATED: diagnostic snapshot
    "FRK_DiagSync"(Index := #Core.RegIndex, Withdraw := FALSE,
        Status := #Status, Held := #Core.Held,
        Timeout := #ParCfg.Timeout, ActiveTimeoutMs := #Core.TimeoutMs);
    // ---- GENERATED: frame end
END_FUNCTION_BLOCK
FUNCTION "FRK_Route_DeclarationUnit" : Bool
{ S7_Optimized_Access := 'TRUE' }
VERSION : 0.1
VAR_INPUT
    Request : "ST_HmiRequest";
END_VAR
VAR_IN_OUT
    Module : "FB_DeclarationUnit";
    Hal : "ST_DeclarationUnitHal";
    Report : "ST_ReleaseReport";
END_VAR
VAR_TEMP
    RouteMatched : Bool;
    Index : Int;
END_VAR
BEGIN
    #FRK_Route_DeclarationUnit := FALSE;
    IF NOT "FRK_PathOwned"(OwnerPath := #Module.Status.Name, TargetPath := #Request.TargetPath) THEN RETURN; END_IF;
    "FRK_Release_DeclarationUnit"(Unit := #Module.Unit, Hal := #Hal);
    "FRK_ManualCommon"(Core := #Module.Core, Unit := #Module.Unit, Status := #Module.Status, Report := #Report);
    IF #Request.TargetPath = STRING_TO_WSTRING(#Module.Status.Name) THEN
        "FRK_ReleaseReason"(Report := #Report, Description := WSTRING#'std.error.unsupportedHmiRequest', Reason := 2008, Path := STRING_TO_WSTRING(#Module.Status.Name), Kind := 4);
        #FRK_Route_DeclarationUnit := TRUE;
        RETURN;
    END_IF;
    #RouteMatched := "FRK_Route_DeclarationCell"(Module := #Module.Cell, Hal := #Hal.Cell, Request := #Request, Report := #Report);
    #FRK_Route_DeclarationUnit := #FRK_Route_DeclarationUnit OR #RouteMatched;
    #RouteMatched := "FRK_Route_SatelliteUnit"(Module := #Module.Satellite, Hal := #Hal.Satellite, Request := #Request, Report := #Report);
    #FRK_Route_DeclarationUnit := #FRK_Route_DeclarationUnit OR #RouteMatched;
END_FUNCTION
FUNCTION "FRK_CfgRestore_DeclarationUnit" : Void
{ S7_Optimized_Access := 'TRUE' }
VERSION : 0.1
VAR_IN_OUT
    Core : "FRK_Core";
    Status : "ST_ModuleStatus";
    ParCfg : "ST_ProductionUnitParCfg";
    StationCfg : "ST_UnitProbeStationCfg";
    ConfigStageParCfg : "ST_ProductionUnitParCfg";
    ConfigDefaultParCfg : "ST_ProductionUnitParCfg";
    ConfigStageStationCfg : "ST_UnitProbeStationCfg";
    ConfigDefaultStationCfg : "ST_UnitProbeStationCfg";
END_VAR
VAR_TEMP
    RootIndex : Int;
    Ok : Bool;
    Stored : Bool;
END_VAR
BEGIN
    #RootIndex := "FRK_ConfigRoot"(RegIndex := #Core.RegIndex);
    IF #RootIndex = 0 THEN RETURN; END_IF;
    #Ok := TRUE;
    #ConfigStageParCfg := #ConfigDefaultParCfg;
    "FRK_CfgDef_DeclarationUnit"(FieldIndex := 1);
    IF "FRK_ConfigFind"(Scope := #Status.Name, Key := "FRK_ConfigScratch".Entry.WriteKey, ModelCode := 'MODEL_A') = 0 THEN
    "FRK_ConfigScratch".Entry.ValueText := DINT_TO_WSTRING(TIME_TO_DINT(#ConfigDefaultParCfg.Timeout));
        #Stored := "FRK_ConfigPut"(Scope := #Status.Name, ModelCode := 'MODEL_A', Text := "FRK_ConfigScratch".Entry.ValueText, RootIndex := #RootIndex);
        IF NOT "FRK_ConfigRuntime".Fresh THEN
            IF "FRK_ConfigStore".ActiveModels[#RootIndex] = 'MODEL_A' THEN #Ok := FALSE; END_IF;
            "FRK_ConfigLoss"(RootIndex := #RootIndex, Scope := #Status.Name);
        END_IF;
    END_IF;
    IF "FRK_ConfigFind"(Scope := #Status.Name, Key := "FRK_ConfigScratch".Entry.WriteKey, ModelCode := 'MODEL_B') = 0 THEN
    "FRK_ConfigScratch".Entry.ValueText := DINT_TO_WSTRING(TIME_TO_DINT(#ConfigDefaultParCfg.Timeout));
        #Stored := "FRK_ConfigPut"(Scope := #Status.Name, ModelCode := 'MODEL_B', Text := "FRK_ConfigScratch".Entry.ValueText, RootIndex := #RootIndex);
        IF NOT "FRK_ConfigRuntime".Fresh THEN
            IF "FRK_ConfigStore".ActiveModels[#RootIndex] = 'MODEL_B' THEN #Ok := FALSE; END_IF;
            "FRK_ConfigLoss"(RootIndex := #RootIndex, Scope := #Status.Name);
        END_IF;
    END_IF;
    #Stored := "FRK_ConfigGet"(Scope := #Status.Name, ModelCode := "FRK_ConfigStore".ActiveModels[#RootIndex]);
    #Ok := #Ok AND #Stored;
    IF #Stored THEN
    #ConfigStageParCfg.Timeout := DINT_TO_TIME(LINT_TO_DINT("FRK_ConfigScratch".Value.Number));
    END_IF;
    "FRK_CfgDef_DeclarationUnit"(FieldIndex := 2);
    IF "FRK_ConfigFind"(Scope := #Status.Name, Key := "FRK_ConfigScratch".Entry.WriteKey, ModelCode := 'MODEL_A') = 0 THEN
    "FRK_ConfigScratch".Entry.ValueText := DINT_TO_WSTRING(#ConfigDefaultParCfg.Preset);
        #Stored := "FRK_ConfigPut"(Scope := #Status.Name, ModelCode := 'MODEL_A', Text := "FRK_ConfigScratch".Entry.ValueText, RootIndex := #RootIndex);
        IF NOT "FRK_ConfigRuntime".Fresh THEN
            IF "FRK_ConfigStore".ActiveModels[#RootIndex] = 'MODEL_A' THEN #Ok := FALSE; END_IF;
            "FRK_ConfigLoss"(RootIndex := #RootIndex, Scope := #Status.Name);
        END_IF;
    END_IF;
    IF "FRK_ConfigFind"(Scope := #Status.Name, Key := "FRK_ConfigScratch".Entry.WriteKey, ModelCode := 'MODEL_B') = 0 THEN
    "FRK_ConfigScratch".Entry.ValueText := DINT_TO_WSTRING(#ConfigDefaultParCfg.Preset);
        #Stored := "FRK_ConfigPut"(Scope := #Status.Name, ModelCode := 'MODEL_B', Text := "FRK_ConfigScratch".Entry.ValueText, RootIndex := #RootIndex);
        IF NOT "FRK_ConfigRuntime".Fresh THEN
            IF "FRK_ConfigStore".ActiveModels[#RootIndex] = 'MODEL_B' THEN #Ok := FALSE; END_IF;
            "FRK_ConfigLoss"(RootIndex := #RootIndex, Scope := #Status.Name);
        END_IF;
    END_IF;
    #Stored := "FRK_ConfigGet"(Scope := #Status.Name, ModelCode := "FRK_ConfigStore".ActiveModels[#RootIndex]);
    #Ok := #Ok AND #Stored;
    IF #Stored THEN
    #ConfigStageParCfg.Preset := LINT_TO_DINT("FRK_ConfigScratch".Value.Number);
    END_IF;
    "FRK_CfgDef_DeclarationUnit"(FieldIndex := 8);
    IF "FRK_ConfigFind"(Scope := #Status.Name, Key := "FRK_ConfigScratch".Entry.WriteKey, ModelCode := 'MODEL_A') = 0 THEN
    "FRK_ConfigScratch".Entry.ValueText := UDINT_TO_WSTRING(#ConfigDefaultParCfg.IdealCycleMs);
        #Stored := "FRK_ConfigPut"(Scope := #Status.Name, ModelCode := 'MODEL_A', Text := "FRK_ConfigScratch".Entry.ValueText, RootIndex := #RootIndex);
        IF NOT "FRK_ConfigRuntime".Fresh THEN
            IF "FRK_ConfigStore".ActiveModels[#RootIndex] = 'MODEL_A' THEN #Ok := FALSE; END_IF;
            "FRK_ConfigLoss"(RootIndex := #RootIndex, Scope := #Status.Name);
        END_IF;
    END_IF;
    IF "FRK_ConfigFind"(Scope := #Status.Name, Key := "FRK_ConfigScratch".Entry.WriteKey, ModelCode := 'MODEL_B') = 0 THEN
    "FRK_ConfigScratch".Entry.ValueText := UDINT_TO_WSTRING(#ConfigDefaultParCfg.IdealCycleMs);
        #Stored := "FRK_ConfigPut"(Scope := #Status.Name, ModelCode := 'MODEL_B', Text := "FRK_ConfigScratch".Entry.ValueText, RootIndex := #RootIndex);
        IF NOT "FRK_ConfigRuntime".Fresh THEN
            IF "FRK_ConfigStore".ActiveModels[#RootIndex] = 'MODEL_B' THEN #Ok := FALSE; END_IF;
            "FRK_ConfigLoss"(RootIndex := #RootIndex, Scope := #Status.Name);
        END_IF;
    END_IF;
    #Stored := "FRK_ConfigGet"(Scope := #Status.Name, ModelCode := "FRK_ConfigStore".ActiveModels[#RootIndex]);
    #Ok := #Ok AND #Stored;
    IF #Stored THEN
    #ConfigStageParCfg.IdealCycleMs := LINT_TO_UDINT("FRK_ConfigScratch".Value.Number);
    END_IF;
    "FRK_CfgDef_DeclarationUnit"(FieldIndex := 9);
    IF "FRK_ConfigFind"(Scope := #Status.Name, Key := "FRK_ConfigScratch".Entry.WriteKey, ModelCode := 'MODEL_A') = 0 THEN
    "FRK_ConfigScratch".Entry.ValueText := UDINT_TO_WSTRING(#ConfigDefaultParCfg.BaselineMs);
        #Stored := "FRK_ConfigPut"(Scope := #Status.Name, ModelCode := 'MODEL_A', Text := "FRK_ConfigScratch".Entry.ValueText, RootIndex := #RootIndex);
        IF NOT "FRK_ConfigRuntime".Fresh THEN
            IF "FRK_ConfigStore".ActiveModels[#RootIndex] = 'MODEL_A' THEN #Ok := FALSE; END_IF;
            "FRK_ConfigLoss"(RootIndex := #RootIndex, Scope := #Status.Name);
        END_IF;
    END_IF;
    IF "FRK_ConfigFind"(Scope := #Status.Name, Key := "FRK_ConfigScratch".Entry.WriteKey, ModelCode := 'MODEL_B') = 0 THEN
    "FRK_ConfigScratch".Entry.ValueText := UDINT_TO_WSTRING(#ConfigDefaultParCfg.BaselineMs);
        #Stored := "FRK_ConfigPut"(Scope := #Status.Name, ModelCode := 'MODEL_B', Text := "FRK_ConfigScratch".Entry.ValueText, RootIndex := #RootIndex);
        IF NOT "FRK_ConfigRuntime".Fresh THEN
            IF "FRK_ConfigStore".ActiveModels[#RootIndex] = 'MODEL_B' THEN #Ok := FALSE; END_IF;
            "FRK_ConfigLoss"(RootIndex := #RootIndex, Scope := #Status.Name);
        END_IF;
    END_IF;
    #Stored := "FRK_ConfigGet"(Scope := #Status.Name, ModelCode := "FRK_ConfigStore".ActiveModels[#RootIndex]);
    #Ok := #Ok AND #Stored;
    IF #Stored THEN
    #ConfigStageParCfg.BaselineMs := LINT_TO_UDINT("FRK_ConfigScratch".Value.Number);
    END_IF;
    IF #Ok THEN
        #ParCfg := #ConfigStageParCfg;
    ELSE
        #ParCfg := #ConfigDefaultParCfg;
        "FRK_ConfigLoss"(RootIndex := #RootIndex, Scope := #Status.Name);
        "FRK_CfgDef_DeclarationUnit"(FieldIndex := 1);
    "FRK_ConfigScratch".Entry.ValueText := DINT_TO_WSTRING(TIME_TO_DINT(#ConfigDefaultParCfg.Timeout));
        #Stored := "FRK_ConfigPut"(Scope := #Status.Name, ModelCode := "FRK_ConfigStore".ActiveModels[#RootIndex], Text := "FRK_ConfigScratch".Entry.ValueText, RootIndex := #RootIndex);
        "FRK_CfgDef_DeclarationUnit"(FieldIndex := 2);
    "FRK_ConfigScratch".Entry.ValueText := DINT_TO_WSTRING(#ConfigDefaultParCfg.Preset);
        #Stored := "FRK_ConfigPut"(Scope := #Status.Name, ModelCode := "FRK_ConfigStore".ActiveModels[#RootIndex], Text := "FRK_ConfigScratch".Entry.ValueText, RootIndex := #RootIndex);
        "FRK_CfgDef_DeclarationUnit"(FieldIndex := 8);
    "FRK_ConfigScratch".Entry.ValueText := UDINT_TO_WSTRING(#ConfigDefaultParCfg.IdealCycleMs);
        #Stored := "FRK_ConfigPut"(Scope := #Status.Name, ModelCode := "FRK_ConfigStore".ActiveModels[#RootIndex], Text := "FRK_ConfigScratch".Entry.ValueText, RootIndex := #RootIndex);
        "FRK_CfgDef_DeclarationUnit"(FieldIndex := 9);
    "FRK_ConfigScratch".Entry.ValueText := UDINT_TO_WSTRING(#ConfigDefaultParCfg.BaselineMs);
        #Stored := "FRK_ConfigPut"(Scope := #Status.Name, ModelCode := "FRK_ConfigStore".ActiveModels[#RootIndex], Text := "FRK_ConfigScratch".Entry.ValueText, RootIndex := #RootIndex);
    END_IF;
    #Ok := TRUE;
    #ConfigStageStationCfg := #ConfigDefaultStationCfg;
    "FRK_CfgDef_DeclarationUnit"(FieldIndex := 3);
    IF "FRK_ConfigFind"(Scope := #Status.Name, Key := "FRK_ConfigScratch".Entry.WriteKey, ModelCode := '') = 0 THEN
    "FRK_ConfigScratch".Entry.ValueText := STRING_TO_WSTRING(#ConfigDefaultStationCfg.SiteLabel);
        #Stored := "FRK_ConfigPut"(Scope := #Status.Name, ModelCode := '', Text := "FRK_ConfigScratch".Entry.ValueText, RootIndex := #RootIndex);
        IF NOT "FRK_ConfigRuntime".Fresh THEN
            #Ok := FALSE;
            "FRK_ConfigLoss"(RootIndex := #RootIndex, Scope := #Status.Name);
        END_IF;
    END_IF;
    #Stored := "FRK_ConfigGet"(Scope := #Status.Name, ModelCode := '');
    #Ok := #Ok AND #Stored;
    IF #Stored THEN
    #ConfigStageStationCfg.SiteLabel := "FRK_ConfigScratch".Value.Text;
    END_IF;
    "FRK_CfgDef_DeclarationUnit"(FieldIndex := 4);
    IF "FRK_ConfigFind"(Scope := #Status.Name, Key := "FRK_ConfigScratch".Entry.WriteKey, ModelCode := '') = 0 THEN
    IF #ConfigDefaultStationCfg.Enabled THEN "FRK_ConfigScratch".Entry.ValueText := WSTRING#'true'; ELSE "FRK_ConfigScratch".Entry.ValueText := WSTRING#'false'; END_IF;
        #Stored := "FRK_ConfigPut"(Scope := #Status.Name, ModelCode := '', Text := "FRK_ConfigScratch".Entry.ValueText, RootIndex := #RootIndex);
        IF NOT "FRK_ConfigRuntime".Fresh THEN
            #Ok := FALSE;
            "FRK_ConfigLoss"(RootIndex := #RootIndex, Scope := #Status.Name);
        END_IF;
    END_IF;
    #Stored := "FRK_ConfigGet"(Scope := #Status.Name, ModelCode := '');
    #Ok := #Ok AND #Stored;
    IF #Stored THEN
    #ConfigStageStationCfg.Enabled := "FRK_ConfigScratch".Value.Flag;
    END_IF;
    "FRK_CfgDef_DeclarationUnit"(FieldIndex := 5);
    IF "FRK_ConfigFind"(Scope := #Status.Name, Key := "FRK_ConfigScratch".Entry.WriteKey, ModelCode := '') = 0 THEN
    "FRK_ConfigScratch".Entry.ValueText := "FRK_ConfigDecimalText"(Number := #ConfigDefaultStationCfg.Ratio);
        #Stored := "FRK_ConfigPut"(Scope := #Status.Name, ModelCode := '', Text := "FRK_ConfigScratch".Entry.ValueText, RootIndex := #RootIndex);
        IF NOT "FRK_ConfigRuntime".Fresh THEN
            #Ok := FALSE;
            "FRK_ConfigLoss"(RootIndex := #RootIndex, Scope := #Status.Name);
        END_IF;
    END_IF;
    #Stored := "FRK_ConfigGet"(Scope := #Status.Name, ModelCode := '');
    #Ok := #Ok AND #Stored;
    IF #Stored THEN
    #ConfigStageStationCfg.Ratio := "FRK_ConfigScratch".Value.Decimal;
    END_IF;
    "FRK_CfgDef_DeclarationUnit"(FieldIndex := 6);
    IF "FRK_ConfigFind"(Scope := #Status.Name, Key := "FRK_ConfigScratch".Entry.WriteKey, ModelCode := '') = 0 THEN
    "FRK_ConfigScratch".Entry.ValueText := "FRK_ConfigDecimalText"(Number := REAL_TO_LREAL(#ConfigDefaultStationCfg.Gain));
        #Stored := "FRK_ConfigPut"(Scope := #Status.Name, ModelCode := '', Text := "FRK_ConfigScratch".Entry.ValueText, RootIndex := #RootIndex);
        IF NOT "FRK_ConfigRuntime".Fresh THEN
            #Ok := FALSE;
            "FRK_ConfigLoss"(RootIndex := #RootIndex, Scope := #Status.Name);
        END_IF;
    END_IF;
    #Stored := "FRK_ConfigGet"(Scope := #Status.Name, ModelCode := '');
    #Ok := #Ok AND #Stored;
    IF #Stored THEN
    #ConfigStageStationCfg.Gain := LREAL_TO_REAL("FRK_ConfigScratch".Value.Decimal);
    END_IF;
    "FRK_CfgDef_DeclarationUnit"(FieldIndex := 7);
    IF "FRK_ConfigFind"(Scope := #Status.Name, Key := "FRK_ConfigScratch".Entry.WriteKey, ModelCode := '') = 0 THEN
    "FRK_ConfigScratch".Entry.ValueText := "FRK_ConfigEnumText"(Number := #ConfigDefaultStationCfg.Grade);
        #Stored := "FRK_ConfigPut"(Scope := #Status.Name, ModelCode := '', Text := "FRK_ConfigScratch".Entry.ValueText, RootIndex := #RootIndex);
        IF NOT "FRK_ConfigRuntime".Fresh THEN
            #Ok := FALSE;
            "FRK_ConfigLoss"(RootIndex := #RootIndex, Scope := #Status.Name);
        END_IF;
    END_IF;
    #Stored := "FRK_ConfigGet"(Scope := #Status.Name, ModelCode := '');
    #Ok := #Ok AND #Stored;
    IF #Stored THEN
    #ConfigStageStationCfg.Grade := LINT_TO_DINT("FRK_ConfigScratch".Value.Number);
    END_IF;
    "FRK_CfgDef_DeclarationUnit"(FieldIndex := 10);
    IF "FRK_ConfigFind"(Scope := #Status.Name, Key := "FRK_ConfigScratch".Entry.WriteKey, ModelCode := '') = 0 THEN
    "FRK_ConfigScratch".Entry.ValueText := UINT_TO_WSTRING(#ConfigDefaultStationCfg.DegradationPercent);
        #Stored := "FRK_ConfigPut"(Scope := #Status.Name, ModelCode := '', Text := "FRK_ConfigScratch".Entry.ValueText, RootIndex := #RootIndex);
        IF NOT "FRK_ConfigRuntime".Fresh THEN
            #Ok := FALSE;
            "FRK_ConfigLoss"(RootIndex := #RootIndex, Scope := #Status.Name);
        END_IF;
    END_IF;
    #Stored := "FRK_ConfigGet"(Scope := #Status.Name, ModelCode := '');
    #Ok := #Ok AND #Stored;
    IF #Stored THEN
    #ConfigStageStationCfg.DegradationPercent := LINT_TO_UINT("FRK_ConfigScratch".Value.Number);
    END_IF;
    "FRK_CfgDef_DeclarationUnit"(FieldIndex := 11);
    IF "FRK_ConfigFind"(Scope := #Status.Name, Key := "FRK_ConfigScratch".Entry.WriteKey, ModelCode := '') = 0 THEN
    "FRK_ConfigScratch".Entry.ValueText := STRING_TO_WSTRING(#ConfigDefaultStationCfg.LongText);
        #Stored := "FRK_ConfigPut"(Scope := #Status.Name, ModelCode := '', Text := "FRK_ConfigScratch".Entry.ValueText, RootIndex := #RootIndex);
        IF NOT "FRK_ConfigRuntime".Fresh THEN
            #Ok := FALSE;
            "FRK_ConfigLoss"(RootIndex := #RootIndex, Scope := #Status.Name);
        END_IF;
    END_IF;
    #Stored := "FRK_ConfigGet"(Scope := #Status.Name, ModelCode := '');
    #Ok := #Ok AND #Stored;
    IF #Stored THEN
    #ConfigStageStationCfg.LongText := "FRK_ConfigScratch".Value.Text;
    END_IF;
    "FRK_CfgDef_DeclarationUnit"(FieldIndex := 12);
    IF "FRK_ConfigFind"(Scope := #Status.Name, Key := "FRK_ConfigScratch".Entry.WriteKey, ModelCode := '') = 0 THEN
    "FRK_ConfigScratch".Entry.ValueText := UDINT_TO_WSTRING(#ConfigDefaultStationCfg.CapturedCycles);
        #Stored := "FRK_ConfigPut"(Scope := #Status.Name, ModelCode := '', Text := "FRK_ConfigScratch".Entry.ValueText, RootIndex := #RootIndex);
        IF NOT "FRK_ConfigRuntime".Fresh THEN
            #Ok := FALSE;
            "FRK_ConfigLoss"(RootIndex := #RootIndex, Scope := #Status.Name);
        END_IF;
    END_IF;
    #Stored := "FRK_ConfigGet"(Scope := #Status.Name, ModelCode := '');
    #Ok := #Ok AND #Stored;
    IF #Stored THEN
    #ConfigStageStationCfg.CapturedCycles := LINT_TO_UDINT("FRK_ConfigScratch".Value.Number);
    END_IF;
    IF #Ok THEN
        #StationCfg := #ConfigStageStationCfg;
    ELSE
        #StationCfg := #ConfigDefaultStationCfg;
        "FRK_ConfigLoss"(RootIndex := #RootIndex, Scope := #Status.Name);
        "FRK_CfgDef_DeclarationUnit"(FieldIndex := 3);
    "FRK_ConfigScratch".Entry.ValueText := STRING_TO_WSTRING(#ConfigDefaultStationCfg.SiteLabel);
        #Stored := "FRK_ConfigPut"(Scope := #Status.Name, ModelCode := '', Text := "FRK_ConfigScratch".Entry.ValueText, RootIndex := #RootIndex);
        "FRK_CfgDef_DeclarationUnit"(FieldIndex := 4);
    IF #ConfigDefaultStationCfg.Enabled THEN "FRK_ConfigScratch".Entry.ValueText := WSTRING#'true'; ELSE "FRK_ConfigScratch".Entry.ValueText := WSTRING#'false'; END_IF;
        #Stored := "FRK_ConfigPut"(Scope := #Status.Name, ModelCode := '', Text := "FRK_ConfigScratch".Entry.ValueText, RootIndex := #RootIndex);
        "FRK_CfgDef_DeclarationUnit"(FieldIndex := 5);
    "FRK_ConfigScratch".Entry.ValueText := "FRK_ConfigDecimalText"(Number := #ConfigDefaultStationCfg.Ratio);
        #Stored := "FRK_ConfigPut"(Scope := #Status.Name, ModelCode := '', Text := "FRK_ConfigScratch".Entry.ValueText, RootIndex := #RootIndex);
        "FRK_CfgDef_DeclarationUnit"(FieldIndex := 6);
    "FRK_ConfigScratch".Entry.ValueText := "FRK_ConfigDecimalText"(Number := REAL_TO_LREAL(#ConfigDefaultStationCfg.Gain));
        #Stored := "FRK_ConfigPut"(Scope := #Status.Name, ModelCode := '', Text := "FRK_ConfigScratch".Entry.ValueText, RootIndex := #RootIndex);
        "FRK_CfgDef_DeclarationUnit"(FieldIndex := 7);
    "FRK_ConfigScratch".Entry.ValueText := "FRK_ConfigEnumText"(Number := #ConfigDefaultStationCfg.Grade);
        #Stored := "FRK_ConfigPut"(Scope := #Status.Name, ModelCode := '', Text := "FRK_ConfigScratch".Entry.ValueText, RootIndex := #RootIndex);
        "FRK_CfgDef_DeclarationUnit"(FieldIndex := 10);
    "FRK_ConfigScratch".Entry.ValueText := UINT_TO_WSTRING(#ConfigDefaultStationCfg.DegradationPercent);
        #Stored := "FRK_ConfigPut"(Scope := #Status.Name, ModelCode := '', Text := "FRK_ConfigScratch".Entry.ValueText, RootIndex := #RootIndex);
        "FRK_CfgDef_DeclarationUnit"(FieldIndex := 11);
    "FRK_ConfigScratch".Entry.ValueText := STRING_TO_WSTRING(#ConfigDefaultStationCfg.LongText);
        #Stored := "FRK_ConfigPut"(Scope := #Status.Name, ModelCode := '', Text := "FRK_ConfigScratch".Entry.ValueText, RootIndex := #RootIndex);
        "FRK_CfgDef_DeclarationUnit"(FieldIndex := 12);
    "FRK_ConfigScratch".Entry.ValueText := UDINT_TO_WSTRING(#ConfigDefaultStationCfg.CapturedCycles);
        #Stored := "FRK_ConfigPut"(Scope := #Status.Name, ModelCode := '', Text := "FRK_ConfigScratch".Entry.ValueText, RootIndex := #RootIndex);
    END_IF;
END_FUNCTION
FUNCTION "FRK_Config_DeclarationUnit" : Void
{ S7_Optimized_Access := 'TRUE' }
VERSION : 0.1
VAR_INPUT
    Access : "FRK_Access";
    RootIndex : Int;
    ModelIndex : UDInt;
END_VAR
VAR_IN_OUT
    Core : "FRK_Core";
    Status : "ST_ModuleStatus";
    ParCfg : "ST_ProductionUnitParCfg";
    ModePolicy : Array[0..6] of "ST_ModePolicy";
    AvailableModelCount : Int;
    ModelCapacity : Int;
    SequenceStepDef : Array[1..8] of "ST_SequenceStepDef";
    SequenceStepCount : Int;
    StationCfg : "ST_UnitProbeStationCfg";
    Cell : "FB_DeclarationCell";
    Satellite : "FB_SatelliteUnit";
    Cursor : "FRK_ConfigCursor";
    Page : "ST_ConfigPage";
END_VAR
VAR_TEMP
    Ok : Bool;
END_VAR
BEGIN
    IF #ModelIndex = 0 THEN
        "FRK_ConfigUnit"(Scope := #Status.Name, Policy := #ModePolicy, ModelCount := #AvailableModelCount, ReadLevel := #Access.Policy.Required[0], Readable := #Access.CurrentLevel >= #Access.Policy.Required[0], Cursor := #Cursor, Page := #Page);
    END_IF;
    IF #ModelIndex = 0 AND #Core.ParentIndex = 0 THEN "FRK_EngineeringManifest"(Scope := #Status.Name, Access := #Access, Cursor := #Cursor, Page := #Page); END_IF;
    IF #ModelIndex = 0 AND #Core.ParentIndex = 0 THEN
        "FRK_ConfigAppend"(Scope := #Status.Name, Item := 'Features/ExportCurrentConfig', ValueText := WSTRING#'true', ValueType := 2, ReadLevel := #Access.Policy.Required[0], Readable := #Access.CurrentLevel >= #Access.Policy.Required[0], Cursor := #Cursor, Page := #Page);
    END_IF;
    IF #ModelIndex = 0 THEN "FRK_ViewManifest"(Scope := #Status.Name, Defs := #SequenceStepDef, Count := #SequenceStepCount, ReadLevel := #Access.Policy.Required[0], Readable := #Access.CurrentLevel >= #Access.Policy.Required[0], Cursor := #Cursor, Page := #Page); END_IF;
    IF #ModelIndex = 0 THEN "FRK_ConfigAppend"(Scope := #Status.Name, Item := 'Features/CaptureConfig', ValueText := WSTRING#'true', ValueType := 2, ReadLevel := #Access.Policy.Required[0], Readable := #Access.CurrentLevel >= #Access.Policy.Required[0], Cursor := #Cursor, Page := #Page); END_IF;
    IF #ModelIndex = 0 THEN
        IF 1 <= #AvailableModelCount THEN "FRK_ConfigAppend"(Scope := #Status.Name, Item := 'AvailableModels/AvailableModels[1]/ModelCode', ValueText := STRING_TO_WSTRING("FRK_ConfigModelCode"(RootIndex := #RootIndex, ModelIndex := 1)), ValueType := 1, ReadLevel := #Access.Policy.Required[0], Readable := #Access.CurrentLevel >= #Access.Policy.Required[0], Cursor := #Cursor, Page := #Page); END_IF;
        IF 2 <= #AvailableModelCount THEN "FRK_ConfigAppend"(Scope := #Status.Name, Item := 'AvailableModels/AvailableModels[2]/ModelCode', ValueText := STRING_TO_WSTRING("FRK_ConfigModelCode"(RootIndex := #RootIndex, ModelIndex := 2)), ValueType := 1, ReadLevel := #Access.Policy.Required[0], Readable := #Access.CurrentLevel >= #Access.Policy.Required[0], Cursor := #Cursor, Page := #Page); END_IF;
        IF 3 <= #AvailableModelCount THEN "FRK_ConfigAppend"(Scope := #Status.Name, Item := 'AvailableModels/AvailableModels[3]/ModelCode', ValueText := STRING_TO_WSTRING("FRK_ConfigModelCode"(RootIndex := #RootIndex, ModelIndex := 3)), ValueType := 1, ReadLevel := #Access.Policy.Required[0], Readable := #Access.CurrentLevel >= #Access.Policy.Required[0], Cursor := #Cursor, Page := #Page); END_IF;
        "FRK_ConfigAppend"(Scope := #Status.Name, Item := 'ModelCapacity', ValueText := INT_TO_WSTRING(#ModelCapacity), ValueType := 0, ReadLevel := #Access.Policy.Required[0], Readable := #Access.CurrentLevel >= #Access.Policy.Required[0], Cursor := #Cursor, Page := #Page);
    END_IF;
    IF (#ModelIndex = 0 OR #Core.ParentIndex = 0) THEN
        "FRK_CfgDef_DeclarationUnit"(FieldIndex := 1);
        "FRK_ConfigScratch".Entry.Scope := STRING_TO_WSTRING(#Status.Name);
        "FRK_ConfigScratch".Entry.ReadLevel := "FRK_DataLevel"(Access := #Access, ClassId := "FRK_ConfigScratch".Entry.ClassId, Minimum := "FRK_ConfigScratch".MinRead, ForWrite := FALSE);
        "FRK_ConfigScratch".Entry.WriteLevel := "FRK_DataLevel"(Access := #Access, ClassId := "FRK_ConfigScratch".Entry.ClassId, Minimum := "FRK_ConfigScratch".MinWrite, ForWrite := TRUE);
        "FRK_ConfigScratch".Entry.Readable := #Access.CurrentLevel >= "FRK_ConfigScratch".Entry.ReadLevel;
        "FRK_ConfigScratch".Entry.ModelScoped := #Core.ParentIndex = 0;
        IF #ModelIndex <> 0 THEN
            "FRK_ConfigScratch".Entry.RequiresReady := "FRK_ConfigScratch".Entry.RequiresReady AND "FRK_ConfigModelCode"(RootIndex := #RootIndex, ModelIndex := #ModelIndex) = "FRK_ConfigStore".ActiveModels[#RootIndex];
            #Ok := "FRK_ConfigGet"(Scope := #Status.Name, ModelCode := "FRK_ConfigModelCode"(RootIndex := #RootIndex, ModelIndex := #ModelIndex));
            IF NOT #Ok THEN "FRK_ConfigScratch".Entry.Readable := FALSE; END_IF;
        ELSE
    "FRK_ConfigScratch".Entry.ValueText := DINT_TO_WSTRING(TIME_TO_DINT(#ParCfg.Timeout));
        END_IF;
        IF NOT "FRK_ConfigScratch".Entry.Readable THEN "FRK_ConfigScratch".Entry.ValueText := WSTRING#''; END_IF;
        "FRK_ConfigAppendEntry"(Cursor := #Cursor, Page := #Page);
    END_IF;
    IF (#ModelIndex = 0 OR #Core.ParentIndex = 0) THEN
        "FRK_CfgDef_DeclarationUnit"(FieldIndex := 2);
        "FRK_ConfigScratch".Entry.Scope := STRING_TO_WSTRING(#Status.Name);
        "FRK_ConfigScratch".Entry.ReadLevel := "FRK_DataLevel"(Access := #Access, ClassId := "FRK_ConfigScratch".Entry.ClassId, Minimum := "FRK_ConfigScratch".MinRead, ForWrite := FALSE);
        "FRK_ConfigScratch".Entry.WriteLevel := "FRK_DataLevel"(Access := #Access, ClassId := "FRK_ConfigScratch".Entry.ClassId, Minimum := "FRK_ConfigScratch".MinWrite, ForWrite := TRUE);
        "FRK_ConfigScratch".Entry.Readable := #Access.CurrentLevel >= "FRK_ConfigScratch".Entry.ReadLevel;
        "FRK_ConfigScratch".Entry.ModelScoped := #Core.ParentIndex = 0;
        IF #ModelIndex <> 0 THEN
            "FRK_ConfigScratch".Entry.RequiresReady := "FRK_ConfigScratch".Entry.RequiresReady AND "FRK_ConfigModelCode"(RootIndex := #RootIndex, ModelIndex := #ModelIndex) = "FRK_ConfigStore".ActiveModels[#RootIndex];
            #Ok := "FRK_ConfigGet"(Scope := #Status.Name, ModelCode := "FRK_ConfigModelCode"(RootIndex := #RootIndex, ModelIndex := #ModelIndex));
            IF NOT #Ok THEN "FRK_ConfigScratch".Entry.Readable := FALSE; END_IF;
        ELSE
    "FRK_ConfigScratch".Entry.ValueText := DINT_TO_WSTRING(#ParCfg.Preset);
        END_IF;
        IF NOT "FRK_ConfigScratch".Entry.Readable THEN "FRK_ConfigScratch".Entry.ValueText := WSTRING#''; END_IF;
        "FRK_ConfigAppendEntry"(Cursor := #Cursor, Page := #Page);
    END_IF;
    IF #ModelIndex = 0 THEN
        "FRK_CfgDef_DeclarationUnit"(FieldIndex := 3);
        "FRK_ConfigScratch".Entry.Scope := STRING_TO_WSTRING(#Status.Name);
        "FRK_ConfigScratch".Entry.ReadLevel := "FRK_DataLevel"(Access := #Access, ClassId := "FRK_ConfigScratch".Entry.ClassId, Minimum := "FRK_ConfigScratch".MinRead, ForWrite := FALSE);
        "FRK_ConfigScratch".Entry.WriteLevel := "FRK_DataLevel"(Access := #Access, ClassId := "FRK_ConfigScratch".Entry.ClassId, Minimum := "FRK_ConfigScratch".MinWrite, ForWrite := TRUE);
        "FRK_ConfigScratch".Entry.Readable := #Access.CurrentLevel >= "FRK_ConfigScratch".Entry.ReadLevel;
        "FRK_ConfigScratch".Entry.ModelScoped := FALSE;
    "FRK_ConfigScratch".Entry.ValueText := STRING_TO_WSTRING(#StationCfg.SiteLabel);
        IF NOT "FRK_ConfigScratch".Entry.Readable THEN "FRK_ConfigScratch".Entry.ValueText := WSTRING#''; END_IF;
        "FRK_ConfigAppendEntry"(Cursor := #Cursor, Page := #Page);
    END_IF;
    IF #ModelIndex = 0 THEN
        "FRK_CfgDef_DeclarationUnit"(FieldIndex := 4);
        "FRK_ConfigScratch".Entry.Scope := STRING_TO_WSTRING(#Status.Name);
        "FRK_ConfigScratch".Entry.ReadLevel := "FRK_DataLevel"(Access := #Access, ClassId := "FRK_ConfigScratch".Entry.ClassId, Minimum := "FRK_ConfigScratch".MinRead, ForWrite := FALSE);
        "FRK_ConfigScratch".Entry.WriteLevel := "FRK_DataLevel"(Access := #Access, ClassId := "FRK_ConfigScratch".Entry.ClassId, Minimum := "FRK_ConfigScratch".MinWrite, ForWrite := TRUE);
        "FRK_ConfigScratch".Entry.Readable := #Access.CurrentLevel >= "FRK_ConfigScratch".Entry.ReadLevel;
        "FRK_ConfigScratch".Entry.ModelScoped := FALSE;
    IF #StationCfg.Enabled THEN "FRK_ConfigScratch".Entry.ValueText := WSTRING#'true'; ELSE "FRK_ConfigScratch".Entry.ValueText := WSTRING#'false'; END_IF;
        IF NOT "FRK_ConfigScratch".Entry.Readable THEN "FRK_ConfigScratch".Entry.ValueText := WSTRING#''; END_IF;
        "FRK_ConfigAppendEntry"(Cursor := #Cursor, Page := #Page);
    END_IF;
    IF #ModelIndex = 0 THEN
        "FRK_CfgDef_DeclarationUnit"(FieldIndex := 5);
        "FRK_ConfigScratch".Entry.Scope := STRING_TO_WSTRING(#Status.Name);
        "FRK_ConfigScratch".Entry.ReadLevel := "FRK_DataLevel"(Access := #Access, ClassId := "FRK_ConfigScratch".Entry.ClassId, Minimum := "FRK_ConfigScratch".MinRead, ForWrite := FALSE);
        "FRK_ConfigScratch".Entry.WriteLevel := "FRK_DataLevel"(Access := #Access, ClassId := "FRK_ConfigScratch".Entry.ClassId, Minimum := "FRK_ConfigScratch".MinWrite, ForWrite := TRUE);
        "FRK_ConfigScratch".Entry.Readable := #Access.CurrentLevel >= "FRK_ConfigScratch".Entry.ReadLevel;
        "FRK_ConfigScratch".Entry.ModelScoped := FALSE;
    "FRK_ConfigScratch".Entry.ValueText := "FRK_ConfigDecimalText"(Number := #StationCfg.Ratio);
        IF "FRK_ConfigScratch".Entry.ValueText = WSTRING#'' THEN "FRK_ConfigScratch".Entry.Readable := FALSE; END_IF;
        IF NOT "FRK_ConfigScratch".Entry.Readable THEN "FRK_ConfigScratch".Entry.ValueText := WSTRING#''; END_IF;
        "FRK_ConfigAppendEntry"(Cursor := #Cursor, Page := #Page);
    END_IF;
    IF #ModelIndex = 0 THEN
        "FRK_CfgDef_DeclarationUnit"(FieldIndex := 6);
        "FRK_ConfigScratch".Entry.Scope := STRING_TO_WSTRING(#Status.Name);
        "FRK_ConfigScratch".Entry.ReadLevel := "FRK_DataLevel"(Access := #Access, ClassId := "FRK_ConfigScratch".Entry.ClassId, Minimum := "FRK_ConfigScratch".MinRead, ForWrite := FALSE);
        "FRK_ConfigScratch".Entry.WriteLevel := "FRK_DataLevel"(Access := #Access, ClassId := "FRK_ConfigScratch".Entry.ClassId, Minimum := "FRK_ConfigScratch".MinWrite, ForWrite := TRUE);
        "FRK_ConfigScratch".Entry.Readable := #Access.CurrentLevel >= "FRK_ConfigScratch".Entry.ReadLevel;
        "FRK_ConfigScratch".Entry.ModelScoped := FALSE;
    "FRK_ConfigScratch".Entry.ValueText := "FRK_ConfigDecimalText"(Number := REAL_TO_LREAL(#StationCfg.Gain));
        IF "FRK_ConfigScratch".Entry.ValueText = WSTRING#'' THEN "FRK_ConfigScratch".Entry.Readable := FALSE; END_IF;
        IF NOT "FRK_ConfigScratch".Entry.Readable THEN "FRK_ConfigScratch".Entry.ValueText := WSTRING#''; END_IF;
        "FRK_ConfigAppendEntry"(Cursor := #Cursor, Page := #Page);
    END_IF;
    IF #ModelIndex = 0 THEN
        "FRK_CfgDef_DeclarationUnit"(FieldIndex := 7);
        "FRK_ConfigScratch".Entry.Scope := STRING_TO_WSTRING(#Status.Name);
        "FRK_ConfigScratch".Entry.ReadLevel := "FRK_DataLevel"(Access := #Access, ClassId := "FRK_ConfigScratch".Entry.ClassId, Minimum := "FRK_ConfigScratch".MinRead, ForWrite := FALSE);
        "FRK_ConfigScratch".Entry.WriteLevel := "FRK_DataLevel"(Access := #Access, ClassId := "FRK_ConfigScratch".Entry.ClassId, Minimum := "FRK_ConfigScratch".MinWrite, ForWrite := TRUE);
        "FRK_ConfigScratch".Entry.Readable := #Access.CurrentLevel >= "FRK_ConfigScratch".Entry.ReadLevel;
        "FRK_ConfigScratch".Entry.ModelScoped := FALSE;
    "FRK_ConfigScratch".Entry.ValueText := "FRK_ConfigEnumText"(Number := #StationCfg.Grade);
        IF NOT "FRK_ConfigScratch".Entry.Readable THEN "FRK_ConfigScratch".Entry.ValueText := WSTRING#''; END_IF;
        "FRK_ConfigAppendEntry"(Cursor := #Cursor, Page := #Page);
    END_IF;
    IF (#ModelIndex = 0 OR #Core.ParentIndex = 0) THEN
        "FRK_CfgDef_DeclarationUnit"(FieldIndex := 8);
        "FRK_ConfigScratch".Entry.Scope := STRING_TO_WSTRING(#Status.Name);
        "FRK_ConfigScratch".Entry.ReadLevel := "FRK_DataLevel"(Access := #Access, ClassId := "FRK_ConfigScratch".Entry.ClassId, Minimum := "FRK_ConfigScratch".MinRead, ForWrite := FALSE);
        "FRK_ConfigScratch".Entry.WriteLevel := "FRK_DataLevel"(Access := #Access, ClassId := "FRK_ConfigScratch".Entry.ClassId, Minimum := "FRK_ConfigScratch".MinWrite, ForWrite := TRUE);
        "FRK_ConfigScratch".Entry.Readable := #Access.CurrentLevel >= "FRK_ConfigScratch".Entry.ReadLevel;
        "FRK_ConfigScratch".Entry.ModelScoped := #Core.ParentIndex = 0;
        IF #ModelIndex <> 0 THEN
            "FRK_ConfigScratch".Entry.RequiresReady := "FRK_ConfigScratch".Entry.RequiresReady AND "FRK_ConfigModelCode"(RootIndex := #RootIndex, ModelIndex := #ModelIndex) = "FRK_ConfigStore".ActiveModels[#RootIndex];
            #Ok := "FRK_ConfigGet"(Scope := #Status.Name, ModelCode := "FRK_ConfigModelCode"(RootIndex := #RootIndex, ModelIndex := #ModelIndex));
            IF NOT #Ok THEN "FRK_ConfigScratch".Entry.Readable := FALSE; END_IF;
        ELSE
    "FRK_ConfigScratch".Entry.ValueText := UDINT_TO_WSTRING(#ParCfg.IdealCycleMs);
        END_IF;
        IF NOT "FRK_ConfigScratch".Entry.Readable THEN "FRK_ConfigScratch".Entry.ValueText := WSTRING#''; END_IF;
        "FRK_ConfigAppendEntry"(Cursor := #Cursor, Page := #Page);
    END_IF;
    IF (#ModelIndex = 0 OR #Core.ParentIndex = 0) THEN
        "FRK_CfgDef_DeclarationUnit"(FieldIndex := 9);
        "FRK_ConfigScratch".Entry.Scope := STRING_TO_WSTRING(#Status.Name);
        "FRK_ConfigScratch".Entry.ReadLevel := "FRK_DataLevel"(Access := #Access, ClassId := "FRK_ConfigScratch".Entry.ClassId, Minimum := "FRK_ConfigScratch".MinRead, ForWrite := FALSE);
        "FRK_ConfigScratch".Entry.WriteLevel := "FRK_DataLevel"(Access := #Access, ClassId := "FRK_ConfigScratch".Entry.ClassId, Minimum := "FRK_ConfigScratch".MinWrite, ForWrite := TRUE);
        "FRK_ConfigScratch".Entry.Readable := #Access.CurrentLevel >= "FRK_ConfigScratch".Entry.ReadLevel;
        "FRK_ConfigScratch".Entry.ModelScoped := #Core.ParentIndex = 0;
        IF #ModelIndex <> 0 THEN
            "FRK_ConfigScratch".Entry.RequiresReady := "FRK_ConfigScratch".Entry.RequiresReady AND "FRK_ConfigModelCode"(RootIndex := #RootIndex, ModelIndex := #ModelIndex) = "FRK_ConfigStore".ActiveModels[#RootIndex];
            #Ok := "FRK_ConfigGet"(Scope := #Status.Name, ModelCode := "FRK_ConfigModelCode"(RootIndex := #RootIndex, ModelIndex := #ModelIndex));
            IF NOT #Ok THEN "FRK_ConfigScratch".Entry.Readable := FALSE; END_IF;
        ELSE
    "FRK_ConfigScratch".Entry.ValueText := UDINT_TO_WSTRING(#ParCfg.BaselineMs);
        END_IF;
        IF NOT "FRK_ConfigScratch".Entry.Readable THEN "FRK_ConfigScratch".Entry.ValueText := WSTRING#''; END_IF;
        "FRK_ConfigAppendEntry"(Cursor := #Cursor, Page := #Page);
    END_IF;
    IF #ModelIndex = 0 THEN
        "FRK_CfgDef_DeclarationUnit"(FieldIndex := 10);
        "FRK_ConfigScratch".Entry.Scope := STRING_TO_WSTRING(#Status.Name);
        "FRK_ConfigScratch".Entry.ReadLevel := "FRK_DataLevel"(Access := #Access, ClassId := "FRK_ConfigScratch".Entry.ClassId, Minimum := "FRK_ConfigScratch".MinRead, ForWrite := FALSE);
        "FRK_ConfigScratch".Entry.WriteLevel := "FRK_DataLevel"(Access := #Access, ClassId := "FRK_ConfigScratch".Entry.ClassId, Minimum := "FRK_ConfigScratch".MinWrite, ForWrite := TRUE);
        "FRK_ConfigScratch".Entry.Readable := #Access.CurrentLevel >= "FRK_ConfigScratch".Entry.ReadLevel;
        "FRK_ConfigScratch".Entry.ModelScoped := FALSE;
    "FRK_ConfigScratch".Entry.ValueText := UINT_TO_WSTRING(#StationCfg.DegradationPercent);
        IF NOT "FRK_ConfigScratch".Entry.Readable THEN "FRK_ConfigScratch".Entry.ValueText := WSTRING#''; END_IF;
        "FRK_ConfigAppendEntry"(Cursor := #Cursor, Page := #Page);
    END_IF;
    IF #ModelIndex = 0 THEN
        "FRK_CfgDef_DeclarationUnit"(FieldIndex := 11);
        "FRK_ConfigScratch".Entry.Scope := STRING_TO_WSTRING(#Status.Name);
        "FRK_ConfigScratch".Entry.ReadLevel := "FRK_DataLevel"(Access := #Access, ClassId := "FRK_ConfigScratch".Entry.ClassId, Minimum := "FRK_ConfigScratch".MinRead, ForWrite := FALSE);
        "FRK_ConfigScratch".Entry.WriteLevel := "FRK_DataLevel"(Access := #Access, ClassId := "FRK_ConfigScratch".Entry.ClassId, Minimum := "FRK_ConfigScratch".MinWrite, ForWrite := TRUE);
        "FRK_ConfigScratch".Entry.Readable := #Access.CurrentLevel >= "FRK_ConfigScratch".Entry.ReadLevel;
        "FRK_ConfigScratch".Entry.ModelScoped := FALSE;
    "FRK_ConfigScratch".Entry.ValueText := STRING_TO_WSTRING(#StationCfg.LongText);
        IF NOT "FRK_ConfigScratch".Entry.Readable THEN "FRK_ConfigScratch".Entry.ValueText := WSTRING#''; END_IF;
        "FRK_ConfigAppendEntry"(Cursor := #Cursor, Page := #Page);
    END_IF;
    IF #ModelIndex = 0 THEN
        "FRK_CfgDef_DeclarationUnit"(FieldIndex := 12);
        "FRK_ConfigScratch".Entry.Scope := STRING_TO_WSTRING(#Status.Name);
        "FRK_ConfigScratch".Entry.ReadLevel := "FRK_DataLevel"(Access := #Access, ClassId := "FRK_ConfigScratch".Entry.ClassId, Minimum := "FRK_ConfigScratch".MinRead, ForWrite := FALSE);
        "FRK_ConfigScratch".Entry.WriteLevel := "FRK_DataLevel"(Access := #Access, ClassId := "FRK_ConfigScratch".Entry.ClassId, Minimum := "FRK_ConfigScratch".MinWrite, ForWrite := TRUE);
        "FRK_ConfigScratch".Entry.Readable := #Access.CurrentLevel >= "FRK_ConfigScratch".Entry.ReadLevel;
        "FRK_ConfigScratch".Entry.ModelScoped := FALSE;
    "FRK_ConfigScratch".Entry.ValueText := UDINT_TO_WSTRING(#StationCfg.CapturedCycles);
        IF NOT "FRK_ConfigScratch".Entry.Readable THEN "FRK_ConfigScratch".Entry.ValueText := WSTRING#''; END_IF;
        "FRK_ConfigAppendEntry"(Cursor := #Cursor, Page := #Page);
    END_IF;
    IF #ModelIndex = 0 THEN "FRK_Config_DeclarationCell"(Module := #Cell, Access := #Access, RootIndex := #RootIndex, ModelIndex := #ModelIndex, Cursor := #Cursor, Page := #Page); END_IF;
    IF #ModelIndex = 0 THEN "FRK_Config_SatelliteUnit"(Module := #Satellite, Access := #Access, RootIndex := #RootIndex, ModelIndex := #ModelIndex, Cursor := #Cursor, Page := #Page); END_IF;
END_FUNCTION
FUNCTION "FRK_CfgWrite_DeclarationUnit" : Bool
{ S7_Optimized_Access := 'TRUE' }
VERSION : 0.1
VAR_INPUT
    Request : "ST_HmiRequest";
    Access : "FRK_Access";
    RootIndex : Int;
    RootReady : Bool;
END_VAR
VAR_IN_OUT
    Core : "FRK_Core";
    Status : "ST_ModuleStatus";
    OutImm : "ST_UnitProbeImm";
    ParCfg : "ST_ProductionUnitParCfg";
    StationCfg : "ST_UnitProbeStationCfg";
    Cell : "FB_DeclarationCell";
    Satellite : "FB_SatelliteUnit";
    Matched : Bool;
END_VAR
VAR_TEMP
    Ok : Bool;
    Code : String[64];
    Inactive : Bool;
    Text : WString[255];
END_VAR
BEGIN
    #FRK_CfgWrite_DeclarationUnit := FALSE;
    IF #Request.TargetPath = STRING_TO_WSTRING(#Status.Name) OR (#Request.TargetPath = WSTRING#'' AND #Core.ParentIndex = 0) THEN
        "FRK_CfgDef_DeclarationUnit"(FieldIndex := 1);
        IF #Request.NameValue = "FRK_ConfigScratch".Entry.WriteKey THEN
            #Matched := TRUE;
            "FRK_ConfigScratch".CommittedScope := #Status.Name;
            IF DINT_TO_UDINT(#Request.IntValue) <> "FRK_ConfigScratch".Entry.WriteRevision THEN RETURN; END_IF;
            IF NOT "FRK_ConfigDataAllowed"(Access := #Access, ForWrite := TRUE, Scope := #Status.Name) THEN
                "FRK_ConfigScratch".RejectDescription := WSTRING#'std.error.accessDenied';
                "FRK_ConfigScratch".RejectReason := 2002; RETURN; END_IF;
            IF #Request.DurationMs <> 0 AND #Core.ParentIndex <> 0 THEN RETURN; END_IF;
            #Code := "FRK_ConfigModelCode"(RootIndex := #RootIndex, ModelIndex := #Request.DurationMs);
            #Inactive := #Code <> "FRK_ConfigStore".ActiveModels[#RootIndex];
            IF "FRK_ConfigScratch".Entry.RequiresReady AND NOT #Inactive AND NOT #RootReady THEN
                "FRK_ConfigScratch".RejectDescription := WSTRING#'std.release.unitNotReady';
                "FRK_ConfigScratch".RejectReason := 2002; RETURN; END_IF;
            #Text := #Request.TextValue;
            IF #Request.Kind = 27 THEN RETURN; END_IF;
            #Ok := "FRK_ConfigPut"(Scope := #Status.Name, ModelCode := #Code, Text := #Text, RootIndex := #RootIndex);
            IF NOT #Ok THEN RETURN; END_IF;
            "FRK_ConfigScratch".CommittedText := #Text; "FRK_ConfigScratch".CommittedScope := #Status.Name;
            IF NOT #Inactive THEN
    #ParCfg.Timeout := DINT_TO_TIME(LINT_TO_DINT("FRK_ConfigScratch".Value.Number));
            END_IF;
            #FRK_CfgWrite_DeclarationUnit := TRUE;
            RETURN;
        END_IF;
        "FRK_CfgDef_DeclarationUnit"(FieldIndex := 2);
        IF #Request.NameValue = "FRK_ConfigScratch".Entry.WriteKey THEN
            #Matched := TRUE;
            "FRK_ConfigScratch".CommittedScope := #Status.Name;
            IF DINT_TO_UDINT(#Request.IntValue) <> "FRK_ConfigScratch".Entry.WriteRevision THEN RETURN; END_IF;
            IF NOT "FRK_ConfigDataAllowed"(Access := #Access, ForWrite := TRUE, Scope := #Status.Name) THEN
                "FRK_ConfigScratch".RejectDescription := WSTRING#'std.error.accessDenied';
                "FRK_ConfigScratch".RejectReason := 2002; RETURN; END_IF;
            IF #Request.DurationMs <> 0 AND #Core.ParentIndex <> 0 THEN RETURN; END_IF;
            #Code := "FRK_ConfigModelCode"(RootIndex := #RootIndex, ModelIndex := #Request.DurationMs);
            #Inactive := #Code <> "FRK_ConfigStore".ActiveModels[#RootIndex];
            IF "FRK_ConfigScratch".Entry.RequiresReady AND NOT #Inactive AND NOT #RootReady THEN
                "FRK_ConfigScratch".RejectDescription := WSTRING#'std.release.unitNotReady';
                "FRK_ConfigScratch".RejectReason := 2002; RETURN; END_IF;
            #Text := #Request.TextValue;
            IF #Request.Kind = 27 THEN RETURN; END_IF;
            #Ok := "FRK_ConfigPut"(Scope := #Status.Name, ModelCode := #Code, Text := #Text, RootIndex := #RootIndex);
            IF NOT #Ok THEN RETURN; END_IF;
            "FRK_ConfigScratch".CommittedText := #Text; "FRK_ConfigScratch".CommittedScope := #Status.Name;
            IF NOT #Inactive THEN
    #ParCfg.Preset := LINT_TO_DINT("FRK_ConfigScratch".Value.Number);
            END_IF;
            #FRK_CfgWrite_DeclarationUnit := TRUE;
            RETURN;
        END_IF;
        "FRK_CfgDef_DeclarationUnit"(FieldIndex := 3);
        IF #Request.NameValue = "FRK_ConfigScratch".Entry.WriteKey THEN
            #Matched := TRUE;
            "FRK_ConfigScratch".CommittedScope := #Status.Name;
            IF DINT_TO_UDINT(#Request.IntValue) <> "FRK_ConfigScratch".Entry.WriteRevision THEN RETURN; END_IF;
            IF NOT "FRK_ConfigDataAllowed"(Access := #Access, ForWrite := TRUE, Scope := #Status.Name) THEN
                "FRK_ConfigScratch".RejectDescription := WSTRING#'std.error.accessDenied';
                "FRK_ConfigScratch".RejectReason := 2002; RETURN; END_IF;
            IF #Request.DurationMs <> 0 THEN RETURN; END_IF;
            #Code := '';
            #Inactive := FALSE;
            IF "FRK_ConfigScratch".Entry.RequiresReady AND NOT #Inactive AND NOT #RootReady THEN
                "FRK_ConfigScratch".RejectDescription := WSTRING#'std.release.unitNotReady';
                "FRK_ConfigScratch".RejectReason := 2002; RETURN; END_IF;
            #Text := #Request.TextValue;
            IF #Request.Kind = 27 THEN RETURN; END_IF;
            #Ok := "FRK_ConfigPut"(Scope := #Status.Name, ModelCode := #Code, Text := #Text, RootIndex := #RootIndex);
            IF NOT #Ok THEN RETURN; END_IF;
            "FRK_ConfigScratch".CommittedText := #Text; "FRK_ConfigScratch".CommittedScope := #Status.Name;
            IF NOT #Inactive THEN
    #StationCfg.SiteLabel := "FRK_ConfigScratch".Value.Text;
            END_IF;
            #FRK_CfgWrite_DeclarationUnit := TRUE;
            RETURN;
        END_IF;
        "FRK_CfgDef_DeclarationUnit"(FieldIndex := 4);
        IF #Request.NameValue = "FRK_ConfigScratch".Entry.WriteKey THEN
            #Matched := TRUE;
            "FRK_ConfigScratch".CommittedScope := #Status.Name;
            IF DINT_TO_UDINT(#Request.IntValue) <> "FRK_ConfigScratch".Entry.WriteRevision THEN RETURN; END_IF;
            IF NOT "FRK_ConfigDataAllowed"(Access := #Access, ForWrite := TRUE, Scope := #Status.Name) THEN
                "FRK_ConfigScratch".RejectDescription := WSTRING#'std.error.accessDenied';
                "FRK_ConfigScratch".RejectReason := 2002; RETURN; END_IF;
            IF #Request.DurationMs <> 0 THEN RETURN; END_IF;
            #Code := '';
            #Inactive := FALSE;
            IF "FRK_ConfigScratch".Entry.RequiresReady AND NOT #Inactive AND NOT #RootReady THEN
                "FRK_ConfigScratch".RejectDescription := WSTRING#'std.release.unitNotReady';
                "FRK_ConfigScratch".RejectReason := 2002; RETURN; END_IF;
            #Text := #Request.TextValue;
            IF #Request.Kind = 27 THEN RETURN; END_IF;
            #Ok := "FRK_ConfigPut"(Scope := #Status.Name, ModelCode := #Code, Text := #Text, RootIndex := #RootIndex);
            IF NOT #Ok THEN RETURN; END_IF;
            "FRK_ConfigScratch".CommittedText := #Text; "FRK_ConfigScratch".CommittedScope := #Status.Name;
            IF NOT #Inactive THEN
    #StationCfg.Enabled := "FRK_ConfigScratch".Value.Flag;
            END_IF;
            #FRK_CfgWrite_DeclarationUnit := TRUE;
            RETURN;
        END_IF;
        "FRK_CfgDef_DeclarationUnit"(FieldIndex := 5);
        IF #Request.NameValue = "FRK_ConfigScratch".Entry.WriteKey THEN
            #Matched := TRUE;
            "FRK_ConfigScratch".CommittedScope := #Status.Name;
            IF DINT_TO_UDINT(#Request.IntValue) <> "FRK_ConfigScratch".Entry.WriteRevision THEN RETURN; END_IF;
            IF NOT "FRK_ConfigDataAllowed"(Access := #Access, ForWrite := TRUE, Scope := #Status.Name) THEN
                "FRK_ConfigScratch".RejectDescription := WSTRING#'std.error.accessDenied';
                "FRK_ConfigScratch".RejectReason := 2002; RETURN; END_IF;
            IF #Request.DurationMs <> 0 THEN RETURN; END_IF;
            #Code := '';
            #Inactive := FALSE;
            IF "FRK_ConfigScratch".Entry.RequiresReady AND NOT #Inactive AND NOT #RootReady THEN
                "FRK_ConfigScratch".RejectDescription := WSTRING#'std.release.unitNotReady';
                "FRK_ConfigScratch".RejectReason := 2002; RETURN; END_IF;
            #Text := #Request.TextValue;
            IF #Request.Kind = 27 THEN RETURN; END_IF;
            #Ok := "FRK_ConfigPut"(Scope := #Status.Name, ModelCode := #Code, Text := #Text, RootIndex := #RootIndex);
            IF NOT #Ok THEN RETURN; END_IF;
            "FRK_ConfigScratch".CommittedText := #Text; "FRK_ConfigScratch".CommittedScope := #Status.Name;
            IF NOT #Inactive THEN
    #StationCfg.Ratio := "FRK_ConfigScratch".Value.Decimal;
            END_IF;
            #FRK_CfgWrite_DeclarationUnit := TRUE;
            RETURN;
        END_IF;
        "FRK_CfgDef_DeclarationUnit"(FieldIndex := 6);
        IF #Request.NameValue = "FRK_ConfigScratch".Entry.WriteKey THEN
            #Matched := TRUE;
            "FRK_ConfigScratch".CommittedScope := #Status.Name;
            IF DINT_TO_UDINT(#Request.IntValue) <> "FRK_ConfigScratch".Entry.WriteRevision THEN RETURN; END_IF;
            IF NOT "FRK_ConfigDataAllowed"(Access := #Access, ForWrite := TRUE, Scope := #Status.Name) THEN
                "FRK_ConfigScratch".RejectDescription := WSTRING#'std.error.accessDenied';
                "FRK_ConfigScratch".RejectReason := 2002; RETURN; END_IF;
            IF #Request.DurationMs <> 0 THEN RETURN; END_IF;
            #Code := '';
            #Inactive := FALSE;
            IF "FRK_ConfigScratch".Entry.RequiresReady AND NOT #Inactive AND NOT #RootReady THEN
                "FRK_ConfigScratch".RejectDescription := WSTRING#'std.release.unitNotReady';
                "FRK_ConfigScratch".RejectReason := 2002; RETURN; END_IF;
            #Text := #Request.TextValue;
            IF #Request.Kind = 27 THEN RETURN; END_IF;
            #Ok := "FRK_ConfigPut"(Scope := #Status.Name, ModelCode := #Code, Text := #Text, RootIndex := #RootIndex);
            IF NOT #Ok THEN RETURN; END_IF;
            "FRK_ConfigScratch".CommittedText := #Text; "FRK_ConfigScratch".CommittedScope := #Status.Name;
            IF NOT #Inactive THEN
    #StationCfg.Gain := LREAL_TO_REAL("FRK_ConfigScratch".Value.Decimal);
            END_IF;
            #FRK_CfgWrite_DeclarationUnit := TRUE;
            RETURN;
        END_IF;
        "FRK_CfgDef_DeclarationUnit"(FieldIndex := 7);
        IF #Request.NameValue = "FRK_ConfigScratch".Entry.WriteKey THEN
            #Matched := TRUE;
            "FRK_ConfigScratch".CommittedScope := #Status.Name;
            IF DINT_TO_UDINT(#Request.IntValue) <> "FRK_ConfigScratch".Entry.WriteRevision THEN RETURN; END_IF;
            IF NOT "FRK_ConfigDataAllowed"(Access := #Access, ForWrite := TRUE, Scope := #Status.Name) THEN
                "FRK_ConfigScratch".RejectDescription := WSTRING#'std.error.accessDenied';
                "FRK_ConfigScratch".RejectReason := 2002; RETURN; END_IF;
            IF #Request.DurationMs <> 0 THEN RETURN; END_IF;
            #Code := '';
            #Inactive := FALSE;
            IF "FRK_ConfigScratch".Entry.RequiresReady AND NOT #Inactive AND NOT #RootReady THEN
                "FRK_ConfigScratch".RejectDescription := WSTRING#'std.release.unitNotReady';
                "FRK_ConfigScratch".RejectReason := 2002; RETURN; END_IF;
            #Text := #Request.TextValue;
            IF #Request.Kind = 27 THEN RETURN; END_IF;
            #Ok := "FRK_ConfigPut"(Scope := #Status.Name, ModelCode := #Code, Text := #Text, RootIndex := #RootIndex);
            IF NOT #Ok THEN RETURN; END_IF;
            "FRK_ConfigScratch".CommittedText := #Text; "FRK_ConfigScratch".CommittedScope := #Status.Name;
            IF NOT #Inactive THEN
    #StationCfg.Grade := LINT_TO_DINT("FRK_ConfigScratch".Value.Number);
            END_IF;
            #FRK_CfgWrite_DeclarationUnit := TRUE;
            RETURN;
        END_IF;
        "FRK_CfgDef_DeclarationUnit"(FieldIndex := 8);
        IF #Request.NameValue = "FRK_ConfigScratch".Entry.WriteKey THEN
            #Matched := TRUE;
            "FRK_ConfigScratch".CommittedScope := #Status.Name;
            IF DINT_TO_UDINT(#Request.IntValue) <> "FRK_ConfigScratch".Entry.WriteRevision THEN RETURN; END_IF;
            IF NOT "FRK_ConfigDataAllowed"(Access := #Access, ForWrite := TRUE, Scope := #Status.Name) THEN
                "FRK_ConfigScratch".RejectDescription := WSTRING#'std.error.accessDenied';
                "FRK_ConfigScratch".RejectReason := 2002; RETURN; END_IF;
            IF #Request.DurationMs <> 0 AND #Core.ParentIndex <> 0 THEN RETURN; END_IF;
            #Code := "FRK_ConfigModelCode"(RootIndex := #RootIndex, ModelIndex := #Request.DurationMs);
            #Inactive := #Code <> "FRK_ConfigStore".ActiveModels[#RootIndex];
            IF "FRK_ConfigScratch".Entry.RequiresReady AND NOT #Inactive AND NOT #RootReady THEN
                "FRK_ConfigScratch".RejectDescription := WSTRING#'std.release.unitNotReady';
                "FRK_ConfigScratch".RejectReason := 2002; RETURN; END_IF;
            #Text := #Request.TextValue;
            IF #Request.Kind = 27 THEN RETURN; END_IF;
            #Ok := "FRK_ConfigPut"(Scope := #Status.Name, ModelCode := #Code, Text := #Text, RootIndex := #RootIndex);
            IF NOT #Ok THEN RETURN; END_IF;
            "FRK_ConfigScratch".CommittedText := #Text; "FRK_ConfigScratch".CommittedScope := #Status.Name;
            IF NOT #Inactive THEN
    #ParCfg.IdealCycleMs := LINT_TO_UDINT("FRK_ConfigScratch".Value.Number);
            END_IF;
            #FRK_CfgWrite_DeclarationUnit := TRUE;
            RETURN;
        END_IF;
        "FRK_CfgDef_DeclarationUnit"(FieldIndex := 9);
        IF #Request.NameValue = "FRK_ConfigScratch".Entry.WriteKey THEN
            #Matched := TRUE;
            "FRK_ConfigScratch".CommittedScope := #Status.Name;
            IF DINT_TO_UDINT(#Request.IntValue) <> "FRK_ConfigScratch".Entry.WriteRevision THEN RETURN; END_IF;
            IF NOT "FRK_ConfigDataAllowed"(Access := #Access, ForWrite := TRUE, Scope := #Status.Name) THEN
                "FRK_ConfigScratch".RejectDescription := WSTRING#'std.error.accessDenied';
                "FRK_ConfigScratch".RejectReason := 2002; RETURN; END_IF;
            IF #Request.DurationMs <> 0 AND #Core.ParentIndex <> 0 THEN RETURN; END_IF;
            #Code := "FRK_ConfigModelCode"(RootIndex := #RootIndex, ModelIndex := #Request.DurationMs);
            #Inactive := #Code <> "FRK_ConfigStore".ActiveModels[#RootIndex];
            IF "FRK_ConfigScratch".Entry.RequiresReady AND NOT #Inactive AND NOT #RootReady THEN
                "FRK_ConfigScratch".RejectDescription := WSTRING#'std.release.unitNotReady';
                "FRK_ConfigScratch".RejectReason := 2002; RETURN; END_IF;
            #Text := #Request.TextValue;
            IF #Request.Kind = 27 THEN RETURN; END_IF;
            #Ok := "FRK_ConfigPut"(Scope := #Status.Name, ModelCode := #Code, Text := #Text, RootIndex := #RootIndex);
            IF NOT #Ok THEN RETURN; END_IF;
            "FRK_ConfigScratch".CommittedText := #Text; "FRK_ConfigScratch".CommittedScope := #Status.Name;
            IF NOT #Inactive THEN
    #ParCfg.BaselineMs := LINT_TO_UDINT("FRK_ConfigScratch".Value.Number);
            END_IF;
            #FRK_CfgWrite_DeclarationUnit := TRUE;
            RETURN;
        END_IF;
        "FRK_CfgDef_DeclarationUnit"(FieldIndex := 10);
        IF #Request.NameValue = "FRK_ConfigScratch".Entry.WriteKey THEN
            #Matched := TRUE;
            "FRK_ConfigScratch".CommittedScope := #Status.Name;
            IF DINT_TO_UDINT(#Request.IntValue) <> "FRK_ConfigScratch".Entry.WriteRevision THEN RETURN; END_IF;
            IF NOT "FRK_ConfigDataAllowed"(Access := #Access, ForWrite := TRUE, Scope := #Status.Name) THEN
                "FRK_ConfigScratch".RejectDescription := WSTRING#'std.error.accessDenied';
                "FRK_ConfigScratch".RejectReason := 2002; RETURN; END_IF;
            IF #Request.DurationMs <> 0 THEN RETURN; END_IF;
            #Code := '';
            #Inactive := FALSE;
            IF "FRK_ConfigScratch".Entry.RequiresReady AND NOT #Inactive AND NOT #RootReady THEN
                "FRK_ConfigScratch".RejectDescription := WSTRING#'std.release.unitNotReady';
                "FRK_ConfigScratch".RejectReason := 2002; RETURN; END_IF;
            #Text := #Request.TextValue;
            IF #Request.Kind = 27 THEN RETURN; END_IF;
            #Ok := "FRK_ConfigPut"(Scope := #Status.Name, ModelCode := #Code, Text := #Text, RootIndex := #RootIndex);
            IF NOT #Ok THEN RETURN; END_IF;
            "FRK_ConfigScratch".CommittedText := #Text; "FRK_ConfigScratch".CommittedScope := #Status.Name;
            IF NOT #Inactive THEN
    #StationCfg.DegradationPercent := LINT_TO_UINT("FRK_ConfigScratch".Value.Number);
            END_IF;
            #FRK_CfgWrite_DeclarationUnit := TRUE;
            RETURN;
        END_IF;
        "FRK_CfgDef_DeclarationUnit"(FieldIndex := 11);
        IF #Request.NameValue = "FRK_ConfigScratch".Entry.WriteKey THEN
            #Matched := TRUE;
            "FRK_ConfigScratch".CommittedScope := #Status.Name;
            IF DINT_TO_UDINT(#Request.IntValue) <> "FRK_ConfigScratch".Entry.WriteRevision THEN RETURN; END_IF;
            IF NOT "FRK_ConfigDataAllowed"(Access := #Access, ForWrite := TRUE, Scope := #Status.Name) THEN
                "FRK_ConfigScratch".RejectDescription := WSTRING#'std.error.accessDenied';
                "FRK_ConfigScratch".RejectReason := 2002; RETURN; END_IF;
            IF #Request.DurationMs <> 0 THEN RETURN; END_IF;
            #Code := '';
            #Inactive := FALSE;
            IF "FRK_ConfigScratch".Entry.RequiresReady AND NOT #Inactive AND NOT #RootReady THEN
                "FRK_ConfigScratch".RejectDescription := WSTRING#'std.release.unitNotReady';
                "FRK_ConfigScratch".RejectReason := 2002; RETURN; END_IF;
            #Text := #Request.TextValue;
            IF #Request.Kind = 27 THEN RETURN; END_IF;
            #Ok := "FRK_ConfigPut"(Scope := #Status.Name, ModelCode := #Code, Text := #Text, RootIndex := #RootIndex);
            IF NOT #Ok THEN RETURN; END_IF;
            "FRK_ConfigScratch".CommittedText := #Text; "FRK_ConfigScratch".CommittedScope := #Status.Name;
            IF NOT #Inactive THEN
    #StationCfg.LongText := "FRK_ConfigScratch".Value.Text;
            END_IF;
            #FRK_CfgWrite_DeclarationUnit := TRUE;
            RETURN;
        END_IF;
        "FRK_CfgDef_DeclarationUnit"(FieldIndex := 12);
        IF #Request.NameValue = "FRK_ConfigScratch".Entry.WriteKey THEN
            #Matched := TRUE;
            "FRK_ConfigScratch".CommittedScope := #Status.Name;
            IF DINT_TO_UDINT(#Request.IntValue) <> "FRK_ConfigScratch".Entry.WriteRevision THEN RETURN; END_IF;
            IF NOT "FRK_ConfigDataAllowed"(Access := #Access, ForWrite := TRUE, Scope := #Status.Name) THEN
                "FRK_ConfigScratch".RejectDescription := WSTRING#'std.error.accessDenied';
                "FRK_ConfigScratch".RejectReason := 2002; RETURN; END_IF;
            IF #Request.DurationMs <> 0 THEN RETURN; END_IF;
            #Code := '';
            #Inactive := FALSE;
            IF "FRK_ConfigScratch".Entry.RequiresReady AND NOT #Inactive AND NOT #RootReady THEN
                "FRK_ConfigScratch".RejectDescription := WSTRING#'std.release.unitNotReady';
                "FRK_ConfigScratch".RejectReason := 2002; RETURN; END_IF;
            #Text := #Request.TextValue;
            IF #Request.Kind = 27 THEN
                IF #Inactive OR NOT #RootReady THEN RETURN; END_IF;
    "FRK_ConfigScratch".Entry.ValueText := UDINT_TO_WSTRING(#OutImm.Cycles);
                #Text := "FRK_ConfigScratch".Entry.ValueText;
            END_IF;
            #Ok := "FRK_ConfigPut"(Scope := #Status.Name, ModelCode := #Code, Text := #Text, RootIndex := #RootIndex);
            IF NOT #Ok THEN RETURN; END_IF;
            "FRK_ConfigScratch".CommittedText := #Text; "FRK_ConfigScratch".CommittedScope := #Status.Name;
            IF NOT #Inactive THEN
    #StationCfg.CapturedCycles := LINT_TO_UDINT("FRK_ConfigScratch".Value.Number);
            END_IF;
            #FRK_CfgWrite_DeclarationUnit := TRUE;
            RETURN;
        END_IF;
    END_IF;
    #Ok := "FRK_CfgWrite_DeclarationCell"(Module := #Cell, Access := #Access, Request := #Request, RootIndex := #RootIndex, RootReady := #RootReady, Matched := #Matched);
    IF #Matched THEN #FRK_CfgWrite_DeclarationUnit := #Ok; RETURN; END_IF;
    #Ok := "FRK_CfgWrite_SatelliteUnit"(Module := #Satellite, Access := #Access, Request := #Request, RootIndex := #RootIndex, RootReady := #RootReady, Matched := #Matched);
    IF #Matched THEN #FRK_CfgWrite_DeclarationUnit := #Ok; RETURN; END_IF;
END_FUNCTION
FUNCTION "FRK_CfgRecipe_DeclarationUnit" : Bool
{ S7_Optimized_Access := 'TRUE' }
VERSION : 0.1
VAR_INPUT
    ModelCode : String;
    Phase : Int;
END_VAR
VAR_IN_OUT
    Status : "ST_ModuleStatus";
    ParCfg : "ST_ProductionUnitParCfg";
    ConfigStaged : Bool;
    ConfigStageParCfg : "ST_ProductionUnitParCfg";
    ConfigDefaultParCfg : "ST_ProductionUnitParCfg";
    Cell : "FB_DeclarationCell";
    Satellite : "FB_SatelliteUnit";
    RejectScope : String;
    RejectKey : String;
END_VAR
VAR_TEMP
    Ok : Bool;
END_VAR
BEGIN
    #FRK_CfgRecipe_DeclarationUnit := TRUE;
    IF #Phase = 1 THEN
        #ConfigStaged := FALSE;
        #ConfigStageParCfg := #ConfigDefaultParCfg;
        "FRK_CfgDef_DeclarationUnit"(FieldIndex := 1);
        #Ok := "FRK_ConfigGet"(Scope := #Status.Name, ModelCode := #ModelCode);
        IF NOT #Ok THEN #RejectScope := #Status.Name; #RejectKey := "FRK_ConfigScratch".Entry.WriteKey; #FRK_CfgRecipe_DeclarationUnit := FALSE; RETURN; END_IF;
    #ConfigStageParCfg.Timeout := DINT_TO_TIME(LINT_TO_DINT("FRK_ConfigScratch".Value.Number));
        "FRK_CfgDef_DeclarationUnit"(FieldIndex := 2);
        #Ok := "FRK_ConfigGet"(Scope := #Status.Name, ModelCode := #ModelCode);
        IF NOT #Ok THEN #RejectScope := #Status.Name; #RejectKey := "FRK_ConfigScratch".Entry.WriteKey; #FRK_CfgRecipe_DeclarationUnit := FALSE; RETURN; END_IF;
    #ConfigStageParCfg.Preset := LINT_TO_DINT("FRK_ConfigScratch".Value.Number);
        "FRK_CfgDef_DeclarationUnit"(FieldIndex := 8);
        #Ok := "FRK_ConfigGet"(Scope := #Status.Name, ModelCode := #ModelCode);
        IF NOT #Ok THEN #RejectScope := #Status.Name; #RejectKey := "FRK_ConfigScratch".Entry.WriteKey; #FRK_CfgRecipe_DeclarationUnit := FALSE; RETURN; END_IF;
    #ConfigStageParCfg.IdealCycleMs := LINT_TO_UDINT("FRK_ConfigScratch".Value.Number);
        "FRK_CfgDef_DeclarationUnit"(FieldIndex := 9);
        #Ok := "FRK_ConfigGet"(Scope := #Status.Name, ModelCode := #ModelCode);
        IF NOT #Ok THEN #RejectScope := #Status.Name; #RejectKey := "FRK_ConfigScratch".Entry.WriteKey; #FRK_CfgRecipe_DeclarationUnit := FALSE; RETURN; END_IF;
    #ConfigStageParCfg.BaselineMs := LINT_TO_UDINT("FRK_ConfigScratch".Value.Number);
        #ConfigStaged := TRUE;
    ELSIF #Phase = 2 THEN
        #ParCfg := #ConfigStageParCfg;
        #ConfigStaged := FALSE;
    ELSE #ConfigStaged := FALSE;
    END_IF;
    #Ok := "FRK_CfgRecipe_DeclarationCell"(Module := #Cell, ModelCode := #ModelCode, Phase := #Phase, RejectScope := #RejectScope, RejectKey := #RejectKey);
    IF NOT #Ok THEN #FRK_CfgRecipe_DeclarationUnit := FALSE; RETURN; END_IF;
    #Ok := "FRK_CfgRecipe_SatelliteUnit"(Module := #Satellite, ModelCode := #ModelCode, Phase := #Phase, RejectScope := #RejectScope, RejectKey := #RejectKey);
    IF NOT #Ok THEN #FRK_CfgRecipe_DeclarationUnit := FALSE; RETURN; END_IF;
END_FUNCTION
FUNCTION "FRK_CfgSetWalk_DeclarationUnit" : Bool
{ S7_Optimized_Access := 'TRUE' }
VERSION : 0.1
VAR_INPUT
    RootIndex : Int;
    Phase : Int;
    Access : "FRK_Access";
    Ready : Bool;
END_VAR
VAR_IN_OUT
    Status : "ST_ModuleStatus";
    ParCfg : "ST_ProductionUnitParCfg";
    StationCfg : "ST_UnitProbeStationCfg";
    ConfigStageParCfg : "ST_ProductionUnitParCfg";
    ConfigStageStationCfg : "ST_UnitProbeStationCfg";
    Cell : "FB_DeclarationCell";
    Satellite : "FB_SatelliteUnit";
END_VAR
VAR_TEMP
    Slot : Int;
    Stored : Int;
    Ok : Bool;
END_VAR
BEGIN
    #FRK_CfgSetWalk_DeclarationUnit := FALSE;
    IF #Phase = 1 THEN #ConfigStageParCfg := #ParCfg; END_IF;
    IF #Phase = 1 THEN #ConfigStageStationCfg := #StationCfg; END_IF;
    IF "FRK_SetRuntime".Work[#RootIndex].Payload.Info.Kind = 0 THEN
        "FRK_CfgDef_DeclarationUnit"(FieldIndex := 1);
        "FRK_SetRuntime".Work[#RootIndex].RejectScope := #Status.Name;
        "FRK_SetRuntime".Work[#RootIndex].RejectKey := "FRK_ConfigScratch".Entry.WriteKey;
        IF #Phase = 0 OR #Phase = 5 THEN
            IF #Phase = 5 AND NOT "FRK_ConfigDataAllowed"(Access := #Access, ForWrite := FALSE, Scope := #Status.Name) THEN RETURN; END_IF;
            IF #Phase = 5 AND (0 <> 0 OR "FRK_SetRuntime".Work[#RootIndex].Payload.Info.ModelCode = "FRK_ConfigStore".ActiveModels[#RootIndex]) THEN
    "FRK_ConfigScratch".Entry.ValueText := DINT_TO_WSTRING(TIME_TO_DINT(#ParCfg.Timeout));
                #Ok := "FRK_ConfigValidate"(Text := "FRK_ConfigScratch".Entry.ValueText);
            ELSE
                #Ok := "FRK_ConfigGet"(Scope := #Status.Name, ModelCode := "FRK_SetRuntime".Work[#RootIndex].Payload.Info.ModelCode);
            END_IF;
            IF NOT #Ok OR "FRK_SetRuntime".Work[#RootIndex].Payload.Info.RecordCount >= 28 THEN RETURN; END_IF;
            #Slot := "FRK_SetRuntime".Work[#RootIndex].Payload.Info.RecordCount + 1;
            "FRK_SetRuntime".Work[#RootIndex].Payload.Records[#Slot].Scope := #Status.Name;
            "FRK_SetRuntime".Work[#RootIndex].Payload.Records[#Slot].WriteKey := "FRK_ConfigScratch".Entry.WriteKey;
            "FRK_SetRuntime".Work[#RootIndex].Payload.Records[#Slot].Revision := "FRK_ConfigScratch".Entry.WriteRevision;
            "FRK_SetRuntime".Work[#RootIndex].Payload.Records[#Slot].Kind := "FRK_ConfigScratch".Entry.ConfigKind;
            "FRK_SetRuntime".Work[#RootIndex].Payload.Records[#Slot].ValueType := "FRK_ConfigScratch".Entry.ValueType;
            "FRK_SetRuntime".Work[#RootIndex].Payload.Records[#Slot].ValueText := WSTRING_TO_STRING("FRK_ConfigScratch".Entry.ValueText);
            "FRK_SetRuntime".Work[#RootIndex].Payload.Info.RecordCount := #Slot;
        ELSIF #Phase = 2 THEN
            #Slot := "FRK_SetRecord"(RootIndex := #RootIndex, Scope := #Status.Name, WriteKey := "FRK_ConfigScratch".Entry.WriteKey);
            #Stored := "FRK_SetRuntime".Work[#RootIndex].Targets[#Slot];
            "FRK_ConfigCommit"(SlotIndex := #Stored, ModelCode := "FRK_SetRuntime".Work[#RootIndex].Payload.Info.ModelCode, Schema := "FRK_ConfigScratch".Schema, Record := "FRK_SetRuntime".Work[#RootIndex].Payload.Records[#Slot]);
        ELSE
            #Slot := "FRK_SetCheck"(RootIndex := #RootIndex, Scope := #Status.Name, Access := #Access, Ready := #Ready, WriteAccess := #Phase <> 3, ReserveTarget := #Phase = 1);
            IF #Slot = 0 THEN RETURN; END_IF;
            IF #Phase = 1 THEN
    #ConfigStageParCfg.Timeout := DINT_TO_TIME(LINT_TO_DINT("FRK_ConfigScratch".Value.Number));
            END_IF;
        END_IF;
    END_IF;
    IF "FRK_SetRuntime".Work[#RootIndex].Payload.Info.Kind = 0 THEN
        "FRK_CfgDef_DeclarationUnit"(FieldIndex := 2);
        "FRK_SetRuntime".Work[#RootIndex].RejectScope := #Status.Name;
        "FRK_SetRuntime".Work[#RootIndex].RejectKey := "FRK_ConfigScratch".Entry.WriteKey;
        IF #Phase = 0 OR #Phase = 5 THEN
            IF #Phase = 5 AND NOT "FRK_ConfigDataAllowed"(Access := #Access, ForWrite := FALSE, Scope := #Status.Name) THEN RETURN; END_IF;
            IF #Phase = 5 AND (0 <> 0 OR "FRK_SetRuntime".Work[#RootIndex].Payload.Info.ModelCode = "FRK_ConfigStore".ActiveModels[#RootIndex]) THEN
    "FRK_ConfigScratch".Entry.ValueText := DINT_TO_WSTRING(#ParCfg.Preset);
                #Ok := "FRK_ConfigValidate"(Text := "FRK_ConfigScratch".Entry.ValueText);
            ELSE
                #Ok := "FRK_ConfigGet"(Scope := #Status.Name, ModelCode := "FRK_SetRuntime".Work[#RootIndex].Payload.Info.ModelCode);
            END_IF;
            IF NOT #Ok OR "FRK_SetRuntime".Work[#RootIndex].Payload.Info.RecordCount >= 28 THEN RETURN; END_IF;
            #Slot := "FRK_SetRuntime".Work[#RootIndex].Payload.Info.RecordCount + 1;
            "FRK_SetRuntime".Work[#RootIndex].Payload.Records[#Slot].Scope := #Status.Name;
            "FRK_SetRuntime".Work[#RootIndex].Payload.Records[#Slot].WriteKey := "FRK_ConfigScratch".Entry.WriteKey;
            "FRK_SetRuntime".Work[#RootIndex].Payload.Records[#Slot].Revision := "FRK_ConfigScratch".Entry.WriteRevision;
            "FRK_SetRuntime".Work[#RootIndex].Payload.Records[#Slot].Kind := "FRK_ConfigScratch".Entry.ConfigKind;
            "FRK_SetRuntime".Work[#RootIndex].Payload.Records[#Slot].ValueType := "FRK_ConfigScratch".Entry.ValueType;
            "FRK_SetRuntime".Work[#RootIndex].Payload.Records[#Slot].ValueText := WSTRING_TO_STRING("FRK_ConfigScratch".Entry.ValueText);
            "FRK_SetRuntime".Work[#RootIndex].Payload.Info.RecordCount := #Slot;
        ELSIF #Phase = 2 THEN
            #Slot := "FRK_SetRecord"(RootIndex := #RootIndex, Scope := #Status.Name, WriteKey := "FRK_ConfigScratch".Entry.WriteKey);
            #Stored := "FRK_SetRuntime".Work[#RootIndex].Targets[#Slot];
            "FRK_ConfigCommit"(SlotIndex := #Stored, ModelCode := "FRK_SetRuntime".Work[#RootIndex].Payload.Info.ModelCode, Schema := "FRK_ConfigScratch".Schema, Record := "FRK_SetRuntime".Work[#RootIndex].Payload.Records[#Slot]);
        ELSE
            #Slot := "FRK_SetCheck"(RootIndex := #RootIndex, Scope := #Status.Name, Access := #Access, Ready := #Ready, WriteAccess := #Phase <> 3, ReserveTarget := #Phase = 1);
            IF #Slot = 0 THEN RETURN; END_IF;
            IF #Phase = 1 THEN
    #ConfigStageParCfg.Preset := LINT_TO_DINT("FRK_ConfigScratch".Value.Number);
            END_IF;
        END_IF;
    END_IF;
    IF "FRK_SetRuntime".Work[#RootIndex].Payload.Info.Kind = 1 THEN
        "FRK_CfgDef_DeclarationUnit"(FieldIndex := 3);
        "FRK_SetRuntime".Work[#RootIndex].RejectScope := #Status.Name;
        "FRK_SetRuntime".Work[#RootIndex].RejectKey := "FRK_ConfigScratch".Entry.WriteKey;
        IF #Phase = 0 OR #Phase = 5 THEN
            IF #Phase = 5 AND NOT "FRK_ConfigDataAllowed"(Access := #Access, ForWrite := FALSE, Scope := #Status.Name) THEN RETURN; END_IF;
            IF #Phase = 5 AND (1 <> 0 OR "FRK_SetRuntime".Work[#RootIndex].Payload.Info.ModelCode = "FRK_ConfigStore".ActiveModels[#RootIndex]) THEN
